(* Logix 5000 project; controller TFF vendor 1 type 14 code 107 rev 33.11; software revision 33.04; part 3 of 38 *)

        [4,3].ScaledMax := 100.0, [4,4].Tag := 'PCV012', [4,4].RawMax := 27648, [4,4].ScaledMax := 100.0, [4,5].Tag := 'SPARE', [4,5].RawMax := 27648, [4,5].ScaledMax := 100.0, [4,6].Tag := 'SPARE', [4,6].RawValue := -6912, [4,6].RawMax := 27648, [4,6].ScaledValue := -25.0, [4,6].ScaledMax := 100.0, [4,7].Tag := 'SPARE', [4,7].RawMax := 27648, [4,7].ScaledMax := 100.0, [4,8].Tag := 'AO#1', [4,8].RawMax := 2047, [4,8].ScaledMax := 100.0, [4,8].EnableCfg := 1, [4,9].Tag := 'AO#2', [4,9].RawMax := 2047, [4,9].ScaledMax := 100.0, [4,9].EnableCfg := 1, [4,10].Tag := 'AO#3', [4,10].RawMax := 2047, [4,10].ScaledMax := 100.0, [4,10].EnableCfg := 1, [4,11].Tag := 'AO#4', [4,11].RawMax := 2047, [4,11].ScaledMax := 100.0, [4,11].EnableCfg := 1, [5,0].Tag := 'SIC001', [5,0].RawMax := 27648, [5,0].ScaledMax := 100.0, [5,0].EnableCfg := 1, [5,1].Tag := 'SIC002', [5,1].RawMax := 27648, [5,1].ScaledMax := 100.0, [5,1].EnableCfg := 1, [5,2].Tag := 'PCV010', [5,2].RawMax := 2047, [5,2].ScaledMax := 100.0, [5,2].EnableCfg := 1, [5,3].Tag := 'PCV011', [5,3].RawMax := 27648, [5,3].ScaledMax := 100.0, [5,4].Tag := 'PCV012', [5,4].RawMax := 27648, [5,4].ScaledMax := 100.0, [5,5].Tag := 'SPARE', [5,5].RawMax := 27648, [5,5].ScaledMax := 100.0, [5,6].Tag := 'SPARE', [5,6].RawValue := -6912, [5,6].RawMax := 27648, [5,6].ScaledValue := -25.0, [5,6].ScaledMax := 100.0, [5,7].Tag := 'SPARE', [5,7].RawMax := 27648, [5,7].ScaledMax := 100.0,
        [5,8].Tag := 'AO#1', [5,8].RawMax := 2047, [5,8].ScaledMax := 100.0, [5,8].EnableCfg := 1, [5,9].Tag := 'AO#2', [5,9].RawMax := 2047, [5,9].ScaledMax := 100.0, [5,9].EnableCfg := 1, [5,10].Tag := 'AO#3', [5,10].RawMax := 2047, [5,10].ScaledMax := 100.0, [5,10].EnableCfg := 1, [5,11].Tag := 'AO#4', [5,11].RawMax := 2047, [5,11].ScaledMax := 100.0, [5,11].EnableCfg := 1);
   AnalogPoint : AnalogInput[50] := ([0].TagName := 'AI201B', [0].OutofRange := 1, [0].RawMin := 5529, [0].RawMax := 27648, [0].RawLowLimit := 5253, [0].RawHighLimit := 27924, [0].FilterActual := 1.0, [0].ScaledMax := 200.0, [0].CurrentValue := -49.993214, [0].RangeMax := 200.0, [0].RangeMaxSave := 200.0, [0].RealCfg := 1, [0].EnableCfg := 1, [0].OverrideCfg := 1, [0].EGU := 'mS/cm', [1].TagName := 'WI201', [1].OutofRange := 1, [1].Address := 1, [1].RawMin := 6553, [1].RawMax := 32767, [1].RawLowLimit := 6225, [1].RawHighLimit := 33095, [1].FilterActual := 1.0, [1].ScaledMax := 2000.0, [1].CurrentValue := -499.94724, [1].RangeMax := 2000.0, [1].RangeMaxSave := 2000.0, [1].RealCfg := 1, [1].EnableCfg := 1, [1].OverrideCfg := 1, [1].EGU := 'kg', [2].TagName := 'FI201', [2].OutofRange := 1, [2].Address := 2, [2].RawMin := 6553, [2].RawMax := 32767, [2].RawValue := 323, [2].RawLowLimit := 6225, [2].RawHighLimit := 33095, [2].FilteredRaw := 323, [2].FilterActual := 1.0, [2].ScaledMax := 100.0, [2].CurrentValue := -23.765926, [2].RangeMax := 100.0, [2].RangeMaxSave := 100.0, [2].RealCfg := 1, [2].EnableCfg := 1, [2].OverrideCfg := 1, [2].EGU := 'Lpm', [3].TagName := 'PCV101', [3].Address := 3, [3].RawMin := 6553, [3].RawMax := 32767, [3].RawValue := 12345, [3].RawLowLimit := 6225, [3].RawHighLimit := 33095, [3].FilteredRaw := 12345, [3].FilterActual := 1.0, [3].ScaledMax := 100.0, [3].CurrentValue := 0.059335444,
        [3].RangeMax := 100.0, [3].RangeMaxSave := 100.0, [3].EnableCfg := 1, [3].EGU := '%Clo', [4].TagName := 'PCV201', [4].Address := 4, [4].RawMin := 6553, [4].RawMax := 32767, [4].RawValue := 17653, [4].RawLowLimit := 6225, [4].RawHighLimit := 33095, [4].FilteredRaw := 17653, [4].FilterActual := 1.0, [4].ScaledMax := 100.0, [4].CurrentValue := 51.80897, [4].RangeMax := 100.0, [4].RangeMaxSave := 100.0, [4].EnableCfg := 1, [4].EGU := '%Opn', [5].TagName := 'PI001', [5].Address := 5, [5].RawMin := 6553, [5].RawMax := 32767, [5].RawValue := 32767, [5].RawLowLimit := 3276, [5].RawHighLimit := 33095, [5].FilteredRaw := 32767, [5].FilterActual := 1.0, [5].ScaledMax := 75.0, [5].CurrentValue := 75.0, [5].RangeMax := 75.0, [5].RangeMaxSave := 75.0, [5].RealCfg := 1, [5].EnableCfg := 1, [5].OverrideCfg := 1, [5].EGU := 'psi', [6].TagName := 'PI101', [6].Address := 6, [6].RawMin := 6553, [6].RawMax := 32767, [6].RawValue := 6576, [6].RawLowLimit := 3276, [6].RawHighLimit := 33095, [6].FilterUser := 50, [6].FilteredRaw := 6575, [6].FilterActual := 0.5, [6].ScaledMax := 75.0, [6].CurrentValue := 0.062943466, [6].RangeMax := 75.0, [6].RangeMaxSave := 75.0, [6].RealCfg := 1, [6].EnableCfg := 1, [6].OverrideCfg := 1, [6].EGU := 'psi', [7].TagName := 'PI201', [7].Address := 7, [7].RawMin := 6553, [7].RawMax := 32767, [7].RawValue := 6561, [7].RawLowLimit := 3276,
        [7].RawHighLimit := 33095, [7].FilteredRaw := 6561, [7].FilterActual := 1.0, [7].ScaledMax := 75.0, [7].CurrentValue := 0.022888534, [7].RangeMax := 75.0, [7].RangeMaxSave := 75.0, [7].RealCfg := 1, [7].EnableCfg := 1, [7].OverrideCfg := 1, [7].EGU := 'psi', [8].TagName := 'PI401', [8].Address := 8, [8].RawMin := 6553, [8].RawMax := 32767, [8].RawValue := 6563, [8].RawLowLimit := 3276, [8].RawHighLimit := 33095, [8].FilteredRaw := 6563, [8].FilterActual := 1.0, [8].ScaledMax := 75.0, [8].CurrentValue := 0.028610667, [8].RangeMax := 75.0, [8].RangeMaxSave := 75.0, [8].RealCfg := 1, [8].EnableCfg := 1, [8].OverrideCfg := 1, [8].EGU := 'psi', [9].TagName := 'AI202', [9].Address := 9, [9].RawMin := 5529, [9].RawMax := 27648, [9].RawLowLimit := 5253, [9].RawHighLimit := 27924, [9].FilterActual := 1.0, [9].ScaledMax := 14.0, [9].RangeMax := 14.0, [9].RangeMaxSave := 14.0, [9].EnableCfg := 1, [9].OverrideCfg := 1, [9].EGU := 'pH', [10].TagName := 'AI201A', [10].OutofRange := 1, [10].Address := 10, [10].RawMin := 5529, [10].RawMax := 27648, [10].RawLowLimit := 5253, [10].RawHighLimit := 27924, [10].FilterActual := 1.0, [10].ScaledMax := 120.0, [10].CurrentValue := -29.99593, [10].RangeMax := 120.0, [10].RangeMaxSave := 120.0, [10].RealCfg := 1, [10].EnableCfg := 1, [10].OverrideCfg := 1, [10].EGU := 'mS/cm', [11].TagName := 'AI203', [11].OutofRange := 1, [11].Address := 11,
        [11].RawMin := 5529, [11].RawMax := 27648, [11].RawLowLimit := 5253, [11].RawHighLimit := 27924, [11].FilterActual := 1.0, [11].ScaledMax := 2.0, [11].CurrentValue := -0.49993217, [11].RangeMax := 2.0, [11].RangeMaxSave := 2.0, [11].RealCfg := 1, [11].EnableCfg := 1, [11].OverrideCfg := 1, [11].EGU := 'AU', [12].TagName := 'AI204', [12].OutofRange := 1, [12].Address := 12, [12].RawMin := 5529, [12].RawMax := 27648, [12].RawLowLimit := 5253, [12].RawHighLimit := 27924, [12].FilterActual := 1.0, [12].ScaledMax := 2.0, [12].CurrentValue := -0.49993217, [12].RangeMax := 2.0, [12].RangeMaxSave := 2.0, [12].RealCfg := 1, [12].EnableCfg := 1, [12].OverrideCfg := 1, [12].EGU := 'AU', [13].TagName := 'TI101', [13].OutofRange := 1, [13].Address := 13, [13].RawMin := 5529, [13].RawMax := 27648, [13].RawLowLimit := 5253, [13].RawHighLimit := 27924, [13].FilterActual := 1.0, [13].ScaledMax := 100.0, [13].CurrentValue := -24.996607, [13].RangeMax := 100.0, [13].RangeMaxSave := 100.0, [13].RealCfg := 1, [13].EnableCfg := 1, [13].OverrideCfg := 1, [13].EGU := '$B0C', [14].TagName := 'MIX101', [14].Address := 14, [14].RawMax := 13824, [14].RawLowLimit := -138, [14].RawHighLimit := 13962, [14].FilterActual := 1.0, [14].ScaledMax := 100.0, [14].RangeMax := 100.0, [14].RangeMaxSave := 100.0, [14].RealCfg := 1, [14].EnableCfg := 1, [14].EGU := '%', [15].TagName := 'WI101', [15].Address := 15, [15].RawMax := 99999,
        [15].RawLowLimit := -1000, [15].RawHighLimit := 100999, [15].FilterActual := 1.0, [15].ScaledMax := 999.99, [15].CurrentValue := -127.832535, [15].EnableCfg := 1, [15].OverrideCfg := 1, [16].TagName := 'AI101', [16].Address := 16, [16].RawMin := 6553, [16].RawMax := 32767, [16].RawLowLimit := 6225, [16].RawHighLimit := 33095, [16].FilterActual := 1.0, [16].ScaledMax := 14.0, [16].RangeMax := 14.0, [16].RangeMaxSave := 14.0, [16].EnableCfg := 1, [16].OverrideCfg := 1, [16].EGU := 'pH', [17].TagName := 'AI104', [17].OutofRange := 1, [17].Address := 17, [17].RawMin := 5529, [17].RawMax := 27648, [17].RawLowLimit := 5253, [17].RawHighLimit := 27924, [17].FilterActual := 1.0, [17].ScaledMax := 200.0, [17].CurrentValue := -49.993214, [17].RangeMax := 200.0, [17].RangeMaxSave := 200.0, [17].RealCfg := 1, [17].OverrideCfg := 1, [17].EGU := 'mS/cm', [18].TagName := 'TCU101', [18].OutofRange := 1, [18].Address := 18, [18].RawMin := 5529, [18].RawMax := 27648, [18].RawLowLimit := 5253, [18].RawHighLimit := 27924, [18].FilterActual := 1.0, [18].ScaledMax := 100.0, [18].CurrentValue := -24.996607, [18].RangeMax := 100.0, [18].RangeMaxSave := 100.0, [18].RealCfg := 1, [18].OverrideCfg := 1, [18].EGU := '$B0C', [19].TagName := 'FI101', [19].Address := 19, [19].RawMin := 6553, [19].RawMax := 32767, [19].RawValue := 6555, [19].RawLowLimit := 6225, [19].RawHighLimit := 33095, [19].FilteredRaw := 6555, [19].FilterActual := 1.0, [19].ScaledMax := 100.0,
        [19].RangeMax := 100.0, [19].RangeMaxSave := 100.0, [19].EnableCfg := 1, [19].OverrideCfg := 1, [19].EGU := 'Lpm', [20].TagName := 'FI401', [20].Address := 20, [20].RawMin := 6553, [20].RawMax := 32767, [20].RawValue := 6550, [20].RawLowLimit := 6225, [20].RawHighLimit := 33095, [20].FilteredRaw := 6550, [20].FilterActual := 1.0, [20].ScaledMax := 100.0, [20].RangeMax := 100.0, [20].RangeMaxSave := 100.0, [20].EnableCfg := 1, [20].OverrideCfg := 1, [20].EGU := 'Lpm', [21].TagName := 'PI601', [21].OutofRange := 1, [21].Address := 21, [21].RawMin := 6553, [21].RawMax := 32767, [21].RawLowLimit := 3276, [21].RawHighLimit := 33095, [21].FilterActual := 1.0, [21].ScaledMax := 138.0, [21].CurrentValue := -34.497368, [21].RangeMax := 138.0, [21].RangeMaxSave := 138.0, [21].RealCfg := 1, [21].EnableCfg := 1, [21].OverrideCfg := 1, [21].EGU := 'mbar', [22].TagName := 'SPARE', [22].OutofRange := 1, [22].Address := 22, [22].RawMin := 5529, [22].RawMax := 27648, [22].RawLowLimit := 5253, [22].RawHighLimit := 27924, [22].FilterActual := 1.0, [22].ScaledMax := 100.0, [22].CurrentValue := -24.996607, [22].RangeMax := 100.0, [22].RangeMaxSave := 100.0, [22].RealCfg := 1, [22].EnableCfg := 1, [22].OverrideCfg := 1, [22].EGU := '$B0C', [23].TagName := 'SPARE', [24].TagName := 'SPARE', [25].TagName := 'SPARE', [26].TagName := 'SPARE', [27].TagName := 'SPARE', [28].TagName := 'AI1', [28].OutofRange := 1, [28].Address := 28,
        [28].RawMin := 6553, [28].RawMax := 32767, [28].RawLowLimit := 6225, [28].RawHighLimit := 33095, [28].FilterActual := 1.0, [28].ScaledMax := 100.0, [28].CurrentValue := -24.998093, [28].RangeMax := 100.0, [28].RangeMaxSave := 100.0, [28].RealCfg := 1, [28].EnableCfg := 1, [28].OverrideCfg := 1, [28].EGU := '%', [29].TagName := 'AI2', [29].OutofRange := 1, [29].Address := 29, [29].RawMin := 6553, [29].RawMax := 32767, [29].RawLowLimit := 6225, [29].RawHighLimit := 33095, [29].FilterActual := 1.0, [29].ScaledMax := 100.0, [29].CurrentValue := -24.998093, [29].RangeMax := 100.0, [29].RangeMaxSave := 100.0, [29].RealCfg := 1, [29].EnableCfg := 1, [29].OverrideCfg := 1, [29].EGU := '%', [30].TagName := 'AI3', [30].OutofRange := 1, [30].Address := 30, [30].RawMin := 6553, [30].RawMax := 32767, [30].RawLowLimit := 6225, [30].RawHighLimit := 33095, [30].FilterActual := 1.0, [30].ScaledMax := 100.0, [30].CurrentValue := -24.998093, [30].RangeMax := 100.0, [30].RangeMaxSave := 100.0, [30].RealCfg := 1, [30].EnableCfg := 1, [30].OverrideCfg := 1, [30].EGU := '%', [31].TagName := 'AI4', [31].OutofRange := 1, [31].Address := 31, [31].RawMin := 6553, [31].RawMax := 32767, [31].RawLowLimit := 6225, [31].RawHighLimit := 33095, [31].FilterActual := 1.0, [31].ScaledMax := 100.0, [31].CurrentValue := -24.998093, [31].RangeMax := 100.0, [31].RangeMaxSave := 100.0, [31].RealCfg := 1, [31].EnableCfg := 1, [31].OverrideCfg := 1,
        [31].EGU := '%', [40].TagName := 'DP', [40].Address := 40, [40].RawMin := 6553, [40].RawMax := 32767, [40].RawLowLimit := 6225, [40].RawHighLimit := 33095, [40].FilterActual := 1.0, [40].ScaledMax := 75.0, [40].CurrentValue := 74.93992, [40].RangeMax := 75.0, [40].RangeMaxSave := 75.0, [40].EnableCfg := 1, [40].OverrideCfg := 1, [40].EGU := 'psi', [41].TagName := 'TMP', [41].Address := 41, [41].RawMin := 6553, [41].RawMax := 32767, [41].RawLowLimit := 6225, [41].RawHighLimit := 33095, [41].FilterActual := 1.0, [41].ScaledMax := 75.0, [41].CurrentValue := 37.49857, [41].RangeMax := 75.0, [41].RangeMaxSave := 75.0, [41].EnableCfg := 1, [41].OverrideCfg := 1, [41].EGU := 'psi', [42].TagName := 'FI003', [42].Address := 42, [42].RawMin := 6553, [42].RawMax := 32767, [42].RawLowLimit := 6225, [42].RawHighLimit := 33095, [42].FilterActual := 1.0, [42].ScaledMax := 120.0, [42].RangeMax := 120.0, [42].RangeMaxSave := 120.0, [42].EnableCfg := 1, [42].OverrideCfg := 1, [42].EGU := 'Lpm', [43].Address := 43, [43].RawMin := 6553, [43].RawMax := 32767, [43].OverrideCfg := 1, [44].TagName := 'LI101', [44].Address := 44, [44].RawMin := 6553, [44].RawMax := 32767, [44].RawLowLimit := 6225, [44].RawHighLimit := 33095, [44].FilterActual := 1.0, [44].ScaledMax := 500.0, [44].CurrentValue := -126.566864, [44].RangeMax := 200.0, [44].RangeMaxSave := 200.0, [44].EnableCfg := 1, [44].OverrideCfg := 1, [45].TagName := 'NWP',
        [45].Address := 45, [45].RawMin := 6553, [45].RawMax := 32767, [45].RawLowLimit := 6225, [45].RawHighLimit := 33095, [45].FilterActual := 1.0, [45].ScaledMax := 999.0, [45].RangeMax := 999.0, [45].RangeMaxSave := 999.0, [45].EnableCfg := 1, [45].EGU := 'L/m$B2/', [46].TagName := 'PERM', [46].Address := 46, [46].RawMin := 6553, [46].RawMax := 32767, [46].RawLowLimit := 6225, [46].RawHighLimit := 33095, [46].FilterActual := 1.0, [46].ScaledMax := 999.0, [46].RangeMax := 999.0, [46].RangeMaxSave := 999.0, [46].EnableCfg := 1, [46].EGU := 'L/m$B2/');   // Analog Input Array
        [19]   // Retentate Flow
        [41]   // Trans-Membrane Pressure
        [28]   // Exchange AI#1
        [0]   // Filtrate Conductivity Cleaning
        [10]   // Filtrate Conductivity Process
        [11]   // Filtrate UV
        [12]   // Filtrate UV
        [13]   // Feed Tank Temperature
        [14]   // Mixer Speed
        [15]   // Feed Tank Weight
        [16]   // Feed Tank pH
        [17]   // Feed Tank Conductivity
        [18]   // TCU Temperature
        [1]   // External Filtrate Weight Scale
        [20]   // Transfer Pump Flow
        [21]   // Feed Tank Pressure
        [22]   // Filtrate Temperature
        [29]   // Exchange AI#2
        [30]   // Exchange AI#3
        [2]   // Filtrate Flow
        [31]   // Exchange AI#4
        [3]   // Retentate Pressure Control Valve Position
        [40]   // Differential Pressure
        [42]   // Feed Flow
        [44]   // Feed Tank volume
        [45]   // Normalized Water Permeability
        [46]   // Membrane Permeability
        [4]   // Filtrate Pressure Control Valve Position
        [5]   // Feed Pressure
        [6]   // Retentate Pressure
        [7]   // Filtrate Pressure
        [8]   // Transfer Pump Pressure
        [9]   // Filtrate pH
   AnalogPoint_Storage : AnalogInput[6,50] := ([0,0].TagName := 'PCV032', [0,0].OutofRange := 1, [0,0].RawMin := 6553, [0,0].RawMax := 32767, [0,0].RawValue := 1, [0,0].RawLowLimit := 6225, [0,0].RawHighLimit := 33095, [0,0].FilteredRaw := 1, [0,0].FilterActual := 1.0, [0,0].ScaledMax := 100.0, [0,0].CurrentValue := -24.994278, [0,0].RangeMax := 100.0, [0,0].RangeMaxSave := 100.0, [0,0].RealCfg := 1, [0,0].EnableCfg := 1, [0,0].OverrideCfg := 1, [0,1].TagName := 'AI201B', [0,1].OutofRange := 1, [0,1].Address := 1, [0,1].RawMin := 5529, [0,1].RawMax := 27648, [0,1].RawLowLimit := 5253, [0,1].RawHighLimit := 27924, [0,1].FilterActual := 1.0, [0,1].ScaledMax := 50.0, [0,1].CurrentValue := -12.498303, [0,1].RangeMax := 50.0, [0,1].RangeMaxSave := 50.0, [0,1].RealCfg := 1, [0,1].EnableCfg := 1, [0,1].OverrideCfg := 1, [0,2].TagName := 'AI201A', [0,2].OutofRange := 1, [0,2].Address := 2, [0,2].RawMin := 5529, [0,2].RawMax := 27648, [0,2].RawLowLimit := 5253, [0,2].RawHighLimit := 27924, [0,2].FilterActual := 1.0, [0,2].ScaledMax := 100.0, [0,2].CurrentValue := -24.996607, [0,2].RangeMax := 100.0, [0,2].RangeMaxSave := 100.0, [0,2].RealCfg := 1, [0,2].EnableCfg := 1, [0,2].OverrideCfg := 1, [0,3].TagName := 'AI202', [0,3].OutofRange := 1, [0,3].Address := 3, [0,3].RawMin := 5529, [0,3].RawMax := 27648, [0,3].RawLowLimit := 5253, [0,3].RawHighLimit := 27924, [0,3].FilterActual := 1.0, [0,3].ScaledMax := 14.0, [0,3].CurrentValue := -3.499525, [0,3].RangeMax := 14.0, [0,3].RangeMaxSave := 14.0, [0,3].RealCfg := 1, [0,3].EnableCfg := 1,
        [0,3].OverrideCfg := 1, [0,4].TagName := 'TI201', [0,4].OutofRange := 1, [0,4].Address := 4, [0,4].RawMin := 5529, [0,4].RawMax := 27648, [0,4].RawLowLimit := 5253, [0,4].RawHighLimit := 27924, [0,4].FilterActual := 1.0, [0,4].ScaledMax := 100.0, [0,4].CurrentValue := -24.996607, [0,4].RangeMax := 100.0, [0,4].RangeMaxSave := 100.0, [0,4].RealCfg := 1, [0,4].EnableCfg := 1, [0,4].OverrideCfg := 1, [0,5].TagName := 'AI203', [0,5].OutofRange := 1, [0,5].Address := 5, [0,5].RawMin := 5529, [0,5].RawMax := 27648, [0,5].RawLowLimit := 5253, [0,5].RawHighLimit := 27924, [0,5].FilterActual := 1.0, [0,5].ScaledMax := 2.0, [0,5].CurrentValue := -0.49993217, [0,5].RangeMax := 2.0, [0,5].RangeMaxSave := 2.0, [0,5].RealCfg := 1, [0,5].EnableCfg := 1, [0,5].OverrideCfg := 1, [0,6].TagName := 'AI204', [0,6].OutofRange := 1, [0,6].Address := 6, [0,6].RawMin := 5529, [0,6].RawMax := 27648, [0,6].RawLowLimit := 5253, [0,6].RawHighLimit := 27924, [0,6].FilterActual := 1.0, [0,6].ScaledMax := 2.0, [0,6].CurrentValue := -0.49993217, [0,6].RangeMax := 2.0, [0,6].RangeMaxSave := 2.0, [0,6].RealCfg := 1, [0,6].EnableCfg := 1, [0,6].OverrideCfg := 1, [0,7].TagName := 'AI102', [0,7].OutofRange := 1, [0,7].Address := 7, [0,7].RawMin := 5529, [0,7].RawMax := 27648, [0,7].RawLowLimit := 5253, [0,7].RawHighLimit := 27924, [0,7].FilterActual := 1.0, [0,7].ScaledMax := 100.0, [0,7].CurrentValue := -24.996607, [0,7].RangeMax := 100.0, [0,7].RangeMaxSave := 100.0, [0,7].RealCfg := 1, [0,7].EnableCfg := 1,
        [0,7].OverrideCfg := 1, [0,8].TagName := 'AI103', [0,8].OutofRange := 1, [0,8].Address := 8, [0,8].RawMin := 5529, [0,8].RawMax := 27648, [0,8].RawLowLimit := 5253, [0,8].RawHighLimit := 27924, [0,8].FilterActual := 1.0, [0,8].ScaledMax := 14.0, [0,8].CurrentValue := -3.499525, [0,8].RangeMax := 14.0, [0,8].RangeMaxSave := 14.0, [0,8].RealCfg := 1, [0,8].EnableCfg := 1, [0,8].OverrideCfg := 1, [0,9].TagName := 'PI003', [0,9].OutofRange := 1, [0,9].Address := 9, [0,9].RawMin := 6553, [0,9].RawMax := 32767, [0,9].RawLowLimit := 6225, [0,9].RawHighLimit := 33095, [0,9].FilterActual := 1.0, [0,9].ScaledMax := 6.0, [0,9].CurrentValue := -1.4998856, [0,9].RangeMax := 6.0, [0,9].RangeMaxSave := 6.0, [0,9].RealCfg := 1, [0,9].EnableCfg := 1, [0,9].OverrideCfg := 1, [0,10].TagName := 'FI001', [0,10].Address := 10, [0,10].RawMin := 5529, [0,10].RawMax := 27648, [0,10].RawLowLimit := 5253, [0,10].RawHighLimit := 27924, [0,10].FilterActual := 1.0, [0,10].ScaledMax := 22.0, [0,10].RangeMax := 22.0, [0,10].RangeMaxSave := 22.0, [0,10].EnableCfg := 1, [0,10].OverrideCfg := 1, [0,11].TagName := 'PI001', [0,11].OutofRange := 1, [0,11].Address := 11, [0,11].RawMin := 6553, [0,11].RawMax := 32767, [0,11].RawLowLimit := 6225, [0,11].RawHighLimit := 33095, [0,11].FilterActual := 1.0, [0,11].ScaledMax := 6.0, [0,11].CurrentValue := -1.4998856, [0,11].RangeMax := 6.0, [0,11].RangeMaxSave := 6.0, [0,11].RealCfg := 1, [0,11].EnableCfg := 1, [0,11].OverrideCfg := 1, [0,12].TagName := 'FI002', [0,12].Address := 12,
        [0,12].RawMin := 5529, [0,12].RawMax := 27648, [0,12].RawLowLimit := 5253, [0,12].RawHighLimit := 27924, [0,12].FilterActual := 1.0, [0,12].ScaledMax := 22.0, [0,12].RangeMax := 22.0, [0,12].RangeMaxSave := 22.0, [0,12].EnableCfg := 1, [0,12].OverrideCfg := 1, [0,13].TagName := 'PI002', [0,13].OutofRange := 1, [0,13].Address := 13, [0,13].RawMin := 6553, [0,13].RawMax := 32767, [0,13].RawLowLimit := 6225, [0,13].RawHighLimit := 33095, [0,13].FilterActual := 1.0, [0,13].ScaledMax := 6.0, [0,13].CurrentValue := -1.4998856, [0,13].RangeMax := 6.0, [0,13].RangeMaxSave := 6.0, [0,13].RealCfg := 1, [0,13].EnableCfg := 1, [0,13].OverrideCfg := 1, [0,14].OutofRange := 1, [0,14].Address := 14, [0,14].RawMin := 5529, [0,14].RawMax := 27648, [0,14].RawLowLimit := 5253, [0,14].RawHighLimit := 27924, [0,14].FilterActual := 1.0, [0,14].ScaledMax := 14.0, [0,14].RangeMax := 14.0, [0,14].RangeMaxSave := 14.0, [0,14].RealCfg := 1, [0,14].OverrideCfg := 1, [0,15].OutofRange := 1, [0,15].Address := 15, [0,15].RawMin := 5529, [0,15].RawMax := 27648, [0,15].RawLowLimit := 5253, [0,15].RawHighLimit := 27924, [0,15].FilterActual := 1.0, [0,15].ScaledMax := 2.0, [0,15].CurrentValue := -0.49993217, [0,15].RangeMax := 2.0, [0,15].RangeMaxSave := 2.0, [0,15].RealCfg := 1, [0,15].OverrideCfg := 1, [0,16].OutofRange := 1, [0,16].Address := 16, [0,16].RawMin := 5529, [0,16].RawMax := 27648, [0,16].RawLowLimit := 5253, [0,16].RawHighLimit := 27924, [0,16].FilterActual := 1.0, [0,16].ScaledMax := 2.0, [0,16].CurrentValue := -0.49993217, [0,16].RangeMax := 2.0,
        [0,16].RangeMaxSave := 2.0, [0,16].RealCfg := 1, [0,16].OverrideCfg := 1, [0,17].OutofRange := 1, [0,17].Address := 17, [0,17].RawMin := 5529, [0,17].RawMax := 27648, [0,17].RawLowLimit := 5253, [0,17].RawHighLimit := 27924, [0,17].FilterActual := 1.0, [0,17].ScaledMin := -1.0, [0,17].ScaledMax := 5.0, [0,17].CurrentValue := -2.4997964, [0,17].RangeMin := -1.0, [0,17].RangeMax := 5.0, [0,17].RangeMinSave := -1.0, [0,17].RangeMaxSave := 5.0, [0,17].RealCfg := 1, [0,17].OverrideCfg := 1, [0,18].OutofRange := 1, [0,18].Address := 18, [0,18].RawMin := 5529, [0,18].RawMax := 27648, [0,18].RawLowLimit := 5253, [0,18].RawHighLimit := 27924, [0,18].FilterActual := 1.0, [0,18].ScaledMin := -1.0, [0,18].ScaledMax := 5.0, [0,18].CurrentValue := -2.4997964, [0,18].RangeMin := -1.0, [0,18].RangeMax := 5.0, [0,18].RangeMinSave := -1.0, [0,18].RangeMaxSave := 5.0, [0,18].RealCfg := 1, [0,18].OverrideCfg := 1, [0,19].OutofRange := 1, [0,19].Address := 19, [0,19].RawMin := 5529, [0,19].RawMax := 27648, [0,19].RawLowLimit := 5253, [0,19].RawHighLimit := 27924, [0,19].FilterActual := 1.0, [0,19].ScaledMin := -1.0, [0,19].ScaledMax := 5.0, [0,19].CurrentValue := -2.4997964, [0,19].RangeMin := -1.0, [0,19].RangeMax := 5.0, [0,19].RangeMinSave := -1.0, [0,19].RangeMaxSave := 5.0, [0,19].RealCfg := 1, [0,19].OverrideCfg := 1, [0,20].OutofRange := 1, [0,20].Address := 20, [0,20].RawMin := 5529, [0,20].RawMax := 27648, [0,20].RawLowLimit := 5253, [0,20].RawHighLimit := 27924, [0,20].FilterActual := 1.0, [0,20].ScaledMax := 100.0, [0,20].CurrentValue := -24.996607,
        [0,20].RangeMax := 100.0, [0,20].RangeMaxSave := 100.0, [0,20].RealCfg := 1, [0,20].OverrideCfg := 1, [0,21].OutofRange := 1, [0,21].Address := 21, [0,21].RawMin := 5529, [0,21].RawMax := 27648, [0,21].RawLowLimit := 5253, [0,21].RawHighLimit := 27924, [0,21].FilterActual := 1.0, [0,21].ScaledMax := 100.0, [0,21].CurrentValue := -24.996607, [0,21].RangeMax := 100.0, [0,21].RangeMaxSave := 100.0, [0,21].RealCfg := 1, [0,21].OverrideCfg := 1, [0,22].TagName := 'SPARE', [0,22].Address := 22, [0,22].RawMin := 5529, [0,22].RawMax := 27648, [0,22].RealCfg := 1, [0,22].OverrideCfg := 1, [0,23].TagName := 'SPARE', [0,23].Address := 23, [0,23].RawMin := 5529, [0,23].RawMax := 27648, [0,23].RealCfg := 1, [0,23].OverrideCfg := 1, [0,24].TagName := 'SPARE', [0,24].Address := 24, [0,24].RawMin := 5529, [0,24].RawMax := 27648, [0,24].RealCfg := 1, [0,24].OverrideCfg := 1, [0,25].TagName := 'SPARE', [0,25].Address := 25, [0,25].RawMin := 5529, [0,25].RawMax := 27648, [0,25].RealCfg := 1, [0,25].OverrideCfg := 1, [0,26].TagName := 'SPARE', [0,26].Address := 26, [0,26].RawMin := 5529, [0,26].RawMax := 27648, [0,26].RealCfg := 1, [0,26].OverrideCfg := 1, [0,27].TagName := 'SPARE', [0,27].Address := 27, [0,27].RawMin := 5529, [0,27].RawMax := 27648, [0,27].RealCfg := 1, [0,27].OverrideCfg := 1, [0,28].TagName := 'AI#1', [0,28].OutofRange := 1, [0,28].Address := 28, [0,28].RawMin := 6553, [0,28].RawMax := 32767, [0,28].RawLowLimit := 6225, [0,28].RawHighLimit := 33095,
        [0,28].FilterActual := 1.0, [0,28].ScaledMax := 100.0, [0,28].CurrentValue := -24.998093, [0,28].RangeMax := 100.0, [0,28].RangeMaxSave := 100.0, [0,28].RealCfg := 1, [0,28].EnableCfg := 1, [0,28].OverrideCfg := 1, [0,29].TagName := 'AI#2', [0,29].OutofRange := 1, [0,29].Address := 29, [0,29].RawMin := 6553, [0,29].RawMax := 32767, [0,29].RawLowLimit := 6225, [0,29].RawHighLimit := 33095, [0,29].FilterActual := 1.0, [0,29].ScaledMax := 100.0, [0,29].CurrentValue := -24.998093, [0,29].RangeMax := 100.0, [0,29].RangeMaxSave := 100.0, [0,29].RealCfg := 1, [0,29].EnableCfg := 1, [0,29].OverrideCfg := 1, [0,30].TagName := 'AI#3', [0,30].OutofRange := 1, [0,30].Address := 30, [0,30].RawMin := 6553, [0,30].RawMax := 32767, [0,30].RawValue := 49, [0,30].RawLowLimit := 6225, [0,30].RawHighLimit := 33095, [0,30].FilteredRaw := 49, [0,30].FilterActual := 1.0, [0,30].ScaledMax := 100.0, [0,30].CurrentValue := -24.811169, [0,30].RangeMax := 100.0, [0,30].RangeMaxSave := 100.0, [0,30].RealCfg := 1, [0,30].EnableCfg := 1, [0,30].OverrideCfg := 1, [0,31].TagName := 'AI#4', [0,31].OutofRange := 1, [0,31].Address := 31, [0,31].RawMin := 6553, [0,31].RawMax := 32767, [0,31].RawValue := 48, [0,31].RawLowLimit := 6225, [0,31].RawHighLimit := 33095, [0,31].FilteredRaw := 48, [0,31].FilterActual := 1.0, [0,31].ScaledMax := 100.0, [0,31].CurrentValue := -24.814985, [0,31].RangeMax := 100.0, [0,31].RangeMaxSave := 100.0, [0,31].RealCfg := 1, [0,31].EnableCfg := 1, [0,31].OverrideCfg := 1, [0,40].TagName := 'FI003', [0,40].Address := 40, [0,40].RawMin := 5529,
        [0,40].RawMax := 27648, [0,40].RawLowLimit := 5253, [0,40].RawHighLimit := 27924, [0,40].FilterActual := 1.0, [0,40].ScaledMax := 44.0, [0,40].RangeMax := 44.0, [0,40].RangeMaxSave := 44.0, [0,40].EnableCfg := 1, [0,40].OverrideCfg := 1, [0,41].TagName := 'LV003', [0,41].Address := 41, [0,41].RawMin := 6553, [0,41].RawMax := 32767, [0,41].RawLowLimit := 6225, [0,41].RawHighLimit := 33095, [0,41].FilterActual := 1.0, [0,41].ScaledMax := 9999.0, [0,41].RangeMax := 9999.0, [0,41].RangeMaxSave := 9999.0, [0,41].EnableCfg := 1, [0,41].OverrideCfg := 1, [0,42].TagName := 'LV001', [0,42].Address := 42, [0,42].RawMin := 6553, [0,42].RawMax := 32767, [0,42].RawLowLimit := 6225, [0,42].RawHighLimit := 33095, [0,42].FilterActual := 1.0, [0,42].ScaledMax := 9999.0, [0,42].RangeMax := 9999.0, [0,42].RangeMaxSave := 9999.0, [0,42].EnableCfg := 1, [0,42].OverrideCfg := 1, [0,43].TagName := 'LV002', [0,43].Address := 43, [0,43].RawMin := 6553, [0,43].RawMax := 32767, [0,43].RawLowLimit := 6225, [0,43].RawHighLimit := 33095, [0,43].FilterActual := 1.0, [0,43].ScaledMax := 9999.0, [0,43].RangeMax := 9999.0, [0,43].RangeMaxSave := 9999.0, [0,43].EnableCfg := 1, [0,43].OverrideCfg := 1, [0,44].Address := 44, [0,44].RawMin := 6553, [0,44].RawMax := 32767, [0,44].RawLowLimit := 6225, [0,44].RawHighLimit := 33095, [0,44].FilterActual := 1.0, [0,44].ScaledMax := 99999.0, [0,44].RangeMax := 99999.0, [0,44].RangeMaxSave := 99999.0, [0,45].Address := 42, [0,45].RawMin := 6553, [0,45].RawMax := 32767, [0,45].RawLowLimit := 6225, [0,45].RawHighLimit := 33095, [0,45].FilterActual := 1.0,
        [0,45].ScaledMin := -1.0, [0,45].ScaledMax := 5.0, [0,45].RangeMin := -1.0, [0,45].RangeMax := 5.0, [0,45].RangeMinSave := -1.0, [0,45].RangeMaxSave := 5.0, [0,45].OverrideCfg := 1, [1,0].TagName := 'PCV032', [1,0].OutofRange := 1, [1,0].RawMin := 6553, [1,0].RawMax := 32767, [1,0].RawValue := 1, [1,0].RawLowLimit := 6225, [1,0].RawHighLimit := 33095, [1,0].FilteredRaw := 1, [1,0].FilterActual := 1.0, [1,0].ScaledMax := 100.0, [1,0].CurrentValue := -24.994278, [1,0].RangeMax := 100.0, [1,0].RangeMaxSave := 100.0, [1,0].RealCfg := 1, [1,0].EnableCfg := 1, [1,0].OverrideCfg := 1, [1,1].TagName := 'AI201B', [1,1].OutofRange := 1, [1,1].Address := 1, [1,1].RawMin := 5529, [1,1].RawMax := 27648, [1,1].RawLowLimit := 5253, [1,1].RawHighLimit := 27924, [1,1].FilterActual := 1.0, [1,1].ScaledMax := 50.0, [1,1].CurrentValue := -12.498303, [1,1].RangeMax := 50.0, [1,1].RangeMaxSave := 50.0, [1,1].RealCfg := 1, [1,1].EnableCfg := 1, [1,1].OverrideCfg := 1, [1,2].TagName := 'AI201A', [1,2].OutofRange := 1, [1,2].Address := 2, [1,2].RawMin := 5529, [1,2].RawMax := 27648, [1,2].RawLowLimit := 5253, [1,2].RawHighLimit := 27924, [1,2].FilterActual := 1.0, [1,2].ScaledMax := 100.0, [1,2].CurrentValue := -24.996607, [1,2].RangeMax := 100.0, [1,2].RangeMaxSave := 100.0, [1,2].RealCfg := 1, [1,2].EnableCfg := 1, [1,2].OverrideCfg := 1, [1,3].TagName := 'AI202', [1,3].OutofRange := 1, [1,3].Address := 3, [1,3].RawMin := 5529, [1,3].RawMax := 27648, [1,3].RawLowLimit := 5253, [1,3].RawHighLimit := 27924,
        [1,3].FilterActual := 1.0, [1,3].ScaledMax := 14.0, [1,3].CurrentValue := -3.499525, [1,3].RangeMax := 14.0, [1,3].RangeMaxSave := 14.0, [1,3].RealCfg := 1, [1,3].EnableCfg := 1, [1,3].OverrideCfg := 1, [1,4].TagName := 'TI201', [1,4].OutofRange := 1, [1,4].Address := 4, [1,4].RawMin := 5529, [1,4].RawMax := 27648, [1,4].RawLowLimit := 5253, [1,4].RawHighLimit := 27924, [1,4].FilterActual := 1.0, [1,4].ScaledMax := 100.0, [1,4].CurrentValue := -24.996607, [1,4].RangeMax := 100.0, [1,4].RangeMaxSave := 100.0, [1,4].RealCfg := 1, [1,4].EnableCfg := 1, [1,4].OverrideCfg := 1, [1,5].TagName := 'AI203', [1,5].OutofRange := 1, [1,5].Address := 5, [1,5].RawMin := 5529, [1,5].RawMax := 27648, [1,5].RawLowLimit := 5253, [1,5].RawHighLimit := 27924, [1,5].FilterActual := 1.0, [1,5].ScaledMax := 2.0, [1,5].CurrentValue := -0.49993217, [1,5].RangeMax := 2.0, [1,5].RangeMaxSave := 2.0, [1,5].RealCfg := 1, [1,5].EnableCfg := 1, [1,5].OverrideCfg := 1, [1,6].TagName := 'AI204', [1,6].OutofRange := 1, [1,6].Address := 6, [1,6].RawMin := 5529, [1,6].RawMax := 27648, [1,6].RawLowLimit := 5253, [1,6].RawHighLimit := 27924, [1,6].FilterActual := 1.0, [1,6].ScaledMax := 2.0, [1,6].CurrentValue := -0.49993217, [1,6].RangeMax := 2.0, [1,6].RangeMaxSave := 2.0, [1,6].RealCfg := 1, [1,6].EnableCfg := 1, [1,6].OverrideCfg := 1, [1,7].TagName := 'AI102', [1,7].OutofRange := 1, [1,7].Address := 7, [1,7].RawMin := 5529, [1,7].RawMax := 27648, [1,7].RawLowLimit := 5253, [1,7].RawHighLimit := 27924,
        [1,7].FilterActual := 1.0, [1,7].ScaledMax := 100.0, [1,7].CurrentValue := -24.996607, [1,7].RangeMax := 100.0, [1,7].RangeMaxSave := 100.0, [1,7].RealCfg := 1, [1,7].EnableCfg := 1, [1,7].OverrideCfg := 1, [1,8].TagName := 'AI103', [1,8].OutofRange := 1, [1,8].Address := 8, [1,8].RawMin := 5529, [1,8].RawMax := 27648, [1,8].RawLowLimit := 5253, [1,8].RawHighLimit := 27924, [1,8].FilterActual := 1.0, [1,8].ScaledMax := 14.0, [1,8].CurrentValue := -3.499525, [1,8].RangeMax := 14.0, [1,8].RangeMaxSave := 14.0, [1,8].RealCfg := 1, [1,8].EnableCfg := 1, [1,8].OverrideCfg := 1, [1,9].TagName := 'PI003', [1,9].OutofRange := 1, [1,9].Address := 9, [1,9].RawMin := 6553, [1,9].RawMax := 32767, [1,9].RawLowLimit := 6225, [1,9].RawHighLimit := 33095, [1,9].FilterActual := 1.0, [1,9].ScaledMax := 6.0, [1,9].CurrentValue := -1.4998856, [1,9].RangeMax := 6.0, [1,9].RangeMaxSave := 6.0, [1,9].RealCfg := 1, [1,9].EnableCfg := 1, [1,9].OverrideCfg := 1, [1,10].TagName := 'FI001', [1,10].Address := 10, [1,10].RawMin := 5529, [1,10].RawMax := 27648, [1,10].RawLowLimit := 5253, [1,10].RawHighLimit := 27924, [1,10].FilterActual := 1.0, [1,10].ScaledMax := 22.0, [1,10].RangeMax := 22.0, [1,10].RangeMaxSave := 22.0, [1,10].EnableCfg := 1, [1,10].OverrideCfg := 1, [1,11].TagName := 'PI001', [1,11].OutofRange := 1, [1,11].Address := 11, [1,11].RawMin := 6553, [1,11].RawMax := 32767, [1,11].RawLowLimit := 6225, [1,11].RawHighLimit := 33095, [1,11].FilterActual := 1.0, [1,11].ScaledMax := 6.0, [1,11].CurrentValue := -1.4998856,
        [1,11].RangeMax := 6.0, [1,11].RangeMaxSave := 6.0, [1,11].RealCfg := 1, [1,11].EnableCfg := 1, [1,11].OverrideCfg := 1, [1,12].TagName := 'FI002', [1,12].Address := 12, [1,12].RawMin := 5529, [1,12].RawMax := 27648, [1,12].RawLowLimit := 5253, [1,12].RawHighLimit := 27924, [1,12].FilterActual := 1.0, [1,12].ScaledMax := 22.0, [1,12].RangeMax := 22.0, [1,12].RangeMaxSave := 22.0, [1,12].EnableCfg := 1, [1,12].OverrideCfg := 1, [1,13].TagName := 'PI002', [1,13].OutofRange := 1, [1,13].Address := 13, [1,13].RawMin := 6553, [1,13].RawMax := 32767, [1,13].RawLowLimit := 6225, [1,13].RawHighLimit := 33095, [1,13].FilterActual := 1.0, [1,13].ScaledMax := 6.0, [1,13].CurrentValue := -1.4998856, [1,13].RangeMax := 6.0, [1,13].RangeMaxSave := 6.0, [1,13].RealCfg := 1, [1,13].EnableCfg := 1, [1,13].OverrideCfg := 1, [1,14].OutofRange := 1, [1,14].Address := 14, [1,14].RawMin := 5529, [1,14].RawMax := 27648, [1,14].RawLowLimit := 5253, [1,14].RawHighLimit := 27924, [1,14].FilterActual := 1.0, [1,14].ScaledMax := 14.0, [1,14].RangeMax := 14.0, [1,14].RangeMaxSave := 14.0, [1,14].RealCfg := 1, [1,14].OverrideCfg := 1, [1,15].OutofRange := 1, [1,15].Address := 15, [1,15].RawMin := 5529, [1,15].RawMax := 27648, [1,15].RawLowLimit := 5253, [1,15].RawHighLimit := 27924, [1,15].FilterActual := 1.0, [1,15].ScaledMax := 2.0, [1,15].CurrentValue := -0.49993217, [1,15].RangeMax := 2.0, [1,15].RangeMaxSave := 2.0, [1,15].RealCfg := 1, [1,15].OverrideCfg := 1, [1,16].OutofRange := 1, [1,16].Address := 16, [1,16].RawMin := 5529,
        [1,16].RawMax := 27648, [1,16].RawLowLimit := 5253, [1,16].RawHighLimit := 27924, [1,16].FilterActual := 1.0, [1,16].ScaledMax := 2.0, [1,16].CurrentValue := -0.49993217, [1,16].RangeMax := 2.0, [1,16].RangeMaxSave := 2.0, [1,16].RealCfg := 1, [1,16].OverrideCfg := 1, [1,17].OutofRange := 1, [1,17].Address := 17, [1,17].RawMin := 5529, [1,17].RawMax := 27648, [1,17].RawLowLimit := 5253, [1,17].RawHighLimit := 27924, [1,17].FilterActual := 1.0, [1,17].ScaledMin := -1.0, [1,17].ScaledMax := 5.0, [1,17].CurrentValue := -2.4997964, [1,17].RangeMin := -1.0, [1,17].RangeMax := 5.0, [1,17].RangeMinSave := -1.0, [1,17].RangeMaxSave := 5.0, [1,17].RealCfg := 1, [1,17].OverrideCfg := 1, [1,18].OutofRange := 1, [1,18].Address := 18, [1,18].RawMin := 5529, [1,18].RawMax := 27648, [1,18].RawLowLimit := 5253, [1,18].RawHighLimit := 27924, [1,18].FilterActual := 1.0, [1,18].ScaledMin := -1.0, [1,18].ScaledMax := 5.0, [1,18].CurrentValue := -2.4997964, [1,18].RangeMin := -1.0, [1,18].RangeMax := 5.0, [1,18].RangeMinSave := -1.0, [1,18].RangeMaxSave := 5.0, [1,18].RealCfg := 1, [1,18].OverrideCfg := 1, [1,19].OutofRange := 1, [1,19].Address := 19, [1,19].RawMin := 5529, [1,19].RawMax := 27648, [1,19].RawLowLimit := 5253, [1,19].RawHighLimit := 27924, [1,19].FilterActual := 1.0, [1,19].ScaledMin := -1.0, [1,19].ScaledMax := 5.0, [1,19].CurrentValue := -2.4997964, [1,19].RangeMin := -1.0, [1,19].RangeMax := 5.0, [1,19].RangeMinSave := -1.0, [1,19].RangeMaxSave := 5.0, [1,19].RealCfg := 1, [1,19].OverrideCfg := 1, [1,20].OutofRange := 1, [1,20].Address := 20,
        [1,20].RawMin := 5529, [1,20].RawMax := 27648, [1,20].RawLowLimit := 5253, [1,20].RawHighLimit := 27924, [1,20].FilterActual := 1.0, [1,20].ScaledMax := 100.0, [1,20].CurrentValue := -24.996607, [1,20].RangeMax := 100.0, [1,20].RangeMaxSave := 100.0, [1,20].RealCfg := 1, [1,20].OverrideCfg := 1, [1,21].OutofRange := 1, [1,21].Address := 21, [1,21].RawMin := 5529, [1,21].RawMax := 27648, [1,21].RawLowLimit := 5253, [1,21].RawHighLimit := 27924, [1,21].FilterActual := 1.0, [1,21].ScaledMax := 100.0, [1,21].CurrentValue := -24.996607, [1,21].RangeMax := 100.0, [1,21].RangeMaxSave := 100.0, [1,21].RealCfg := 1, [1,21].OverrideCfg := 1, [1,22].TagName := 'SPARE', [1,22].Address := 22, [1,22].RawMin := 5529, [1,22].RawMax := 27648, [1,22].RealCfg := 1, [1,22].OverrideCfg := 1, [1,23].TagName := 'SPARE', [1,23].Address := 23, [1,23].RawMin := 5529, [1,23].RawMax := 27648, [1,23].RealCfg := 1, [1,23].OverrideCfg := 1, [1,24].TagName := 'SPARE', [1,24].Address := 24, [1,24].RawMin := 5529, [1,24].RawMax := 27648, [1,24].RealCfg := 1, [1,24].OverrideCfg := 1, [1,25].TagName := 'SPARE', [1,25].Address := 25, [1,25].RawMin := 5529, [1,25].RawMax := 27648, [1,25].RealCfg := 1, [1,25].OverrideCfg := 1, [1,26].TagName := 'SPARE', [1,26].Address := 26, [1,26].RawMin := 5529, [1,26].RawMax := 27648, [1,26].RealCfg := 1, [1,26].OverrideCfg := 1, [1,27].TagName := 'SPARE', [1,27].Address := 27, [1,27].RawMin := 5529, [1,27].RawMax := 27648, [1,27].RealCfg := 1, [1,27].OverrideCfg := 1,
        [1,28].TagName := 'AI#1', [1,28].OutofRange := 1, [1,28].Address := 28, [1,28].RawMin := 6553, [1,28].RawMax := 32767, [1,28].RawLowLimit := 6225, [1,28].RawHighLimit := 33095, [1,28].FilterActual := 1.0, [1,28].ScaledMax := 100.0, [1,28].CurrentValue := -24.998093, [1,28].RangeMax := 100.0, [1,28].RangeMaxSave := 100.0, [1,28].RealCfg := 1, [1,28].EnableCfg := 1, [1,28].OverrideCfg := 1, [1,29].TagName := 'AI#2', [1,29].OutofRange := 1, [1,29].Address := 29, [1,29].RawMin := 6553, [1,29].RawMax := 32767, [1,29].RawLowLimit := 6225, [1,29].RawHighLimit := 33095, [1,29].FilterActual := 1.0, [1,29].ScaledMax := 100.0, [1,29].CurrentValue := -24.998093, [1,29].RangeMax := 100.0, [1,29].RangeMaxSave := 100.0, [1,29].RealCfg := 1, [1,29].EnableCfg := 1, [1,29].OverrideCfg := 1, [1,30].TagName := 'AI#3', [1,30].OutofRange := 1, [1,30].Address := 30, [1,30].RawMin := 6553, [1,30].RawMax := 32767, [1,30].RawValue := 49, [1,30].RawLowLimit := 6225, [1,30].RawHighLimit := 33095, [1,30].FilteredRaw := 49, [1,30].FilterActual := 1.0, [1,30].ScaledMax := 100.0, [1,30].CurrentValue := -24.811169, [1,30].RangeMax := 100.0, [1,30].RangeMaxSave := 100.0, [1,30].RealCfg := 1, [1,30].EnableCfg := 1, [1,30].OverrideCfg := 1, [1,31].TagName := 'AI#4', [1,31].OutofRange := 1, [1,31].Address := 31, [1,31].RawMin := 6553, [1,31].RawMax := 32767, [1,31].RawValue := 48, [1,31].RawLowLimit := 6225, [1,31].RawHighLimit := 33095, [1,31].FilteredRaw := 48, [1,31].FilterActual := 1.0, [1,31].ScaledMax := 100.0, [1,31].CurrentValue := -24.814985, [1,31].RangeMax := 100.0,
        [1,31].RangeMaxSave := 100.0, [1,31].RealCfg := 1, [1,31].EnableCfg := 1, [1,31].OverrideCfg := 1, [1,40].TagName := 'FI003', [1,40].Address := 40, [1,40].RawMin := 5529, [1,40].RawMax := 27648, [1,40].RawLowLimit := 5253, [1,40].RawHighLimit := 27924, [1,40].FilterActual := 1.0, [1,40].ScaledMax := 44.0, [1,40].RangeMax := 44.0, [1,40].RangeMaxSave := 44.0, [1,40].EnableCfg := 1, [1,40].OverrideCfg := 1, [1,41].TagName := 'LV003', [1,41].Address := 41, [1,41].RawMin := 6553, [1,41].RawMax := 32767, [1,41].RawLowLimit := 6225, [1,41].RawHighLimit := 33095, [1,41].FilterActual := 1.0, [1,41].ScaledMax := 9999.0, [1,41].RangeMax := 9999.0, [1,41].RangeMaxSave := 9999.0, [1,41].EnableCfg := 1, [1,41].OverrideCfg := 1, [1,42].TagName := 'LV001', [1,42].Address := 42, [1,42].RawMin := 6553, [1,42].RawMax := 32767, [1,42].RawLowLimit := 6225, [1,42].RawHighLimit := 33095, [1,42].FilterActual := 1.0, [1,42].ScaledMax := 9999.0, [1,42].RangeMax := 9999.0, [1,42].RangeMaxSave := 9999.0, [1,42].EnableCfg := 1, [1,42].OverrideCfg := 1, [1,43].TagName := 'LV002', [1,43].Address := 43, [1,43].RawMin := 6553, [1,43].RawMax := 32767, [1,43].RawLowLimit := 6225, [1,43].RawHighLimit := 33095, [1,43].FilterActual := 1.0, [1,43].ScaledMax := 9999.0, [1,43].RangeMax := 9999.0, [1,43].RangeMaxSave := 9999.0, [1,43].EnableCfg := 1, [1,43].OverrideCfg := 1, [1,44].Address := 44, [1,44].RawMin := 6553, [1,44].RawMax := 32767, [1,44].RawLowLimit := 6225, [1,44].RawHighLimit := 33095, [1,44].FilterActual := 1.0, [1,44].ScaledMax := 99999.0, [1,44].RangeMax := 99999.0,
        [1,44].RangeMaxSave := 99999.0, [1,45].Address := 42, [1,45].RawMin := 6553, [1,45].RawMax := 32767, [1,45].RawLowLimit := 6225, [1,45].RawHighLimit := 33095, [1,45].FilterActual := 1.0, [1,45].ScaledMin := -1.0, [1,45].ScaledMax := 5.0, [1,45].RangeMin := -1.0, [1,45].RangeMax := 5.0, [1,45].RangeMinSave := -1.0, [1,45].RangeMaxSave := 5.0, [1,45].OverrideCfg := 1, [2,0].TagName := 'PCV032', [2,0].OutofRange := 1, [2,0].RawMin := 6553, [2,0].RawMax := 32767, [2,0].RawValue := 1, [2,0].RawLowLimit := 6225, [2,0].RawHighLimit := 33095, [2,0].FilteredRaw := 1, [2,0].FilterActual := 1.0, [2,0].ScaledMax := 100.0, [2,0].CurrentValue := -24.994278, [2,0].RangeMax := 100.0, [2,0].RangeMaxSave := 100.0, [2,0].RealCfg := 1, [2,0].EnableCfg := 1, [2,0].OverrideCfg := 1, [2,1].TagName := 'AI201B', [2,1].OutofRange := 1, [2,1].Address := 1, [2,1].RawMin := 5529, [2,1].RawMax := 27648, [2,1].RawLowLimit := 5253, [2,1].RawHighLimit := 27924, [2,1].FilterActual := 1.0, [2,1].ScaledMax := 50.0, [2,1].CurrentValue := -12.498303, [2,1].RangeMax := 50.0, [2,1].RangeMaxSave := 50.0, [2,1].RealCfg := 1, [2,1].EnableCfg := 1, [2,1].OverrideCfg := 1, [2,2].TagName := 'AI201A', [2,2].OutofRange := 1, [2,2].Address := 2, [2,2].RawMin := 5529, [2,2].RawMax := 27648, [2,2].RawLowLimit := 5253, [2,2].RawHighLimit := 27924, [2,2].FilterActual := 1.0, [2,2].ScaledMax := 100.0, [2,2].CurrentValue := -24.996607, [2,2].RangeMax := 100.0, [2,2].RangeMaxSave := 100.0, [2,2].RealCfg := 1, [2,2].EnableCfg := 1, [2,2].OverrideCfg := 1,
        [2,3].TagName := 'AI202', [2,3].OutofRange := 1, [2,3].Address := 3, [2,3].RawMin := 5529, [2,3].RawMax := 27648, [2,3].RawLowLimit := 5253, [2,3].RawHighLimit := 27924, [2,3].FilterActual := 1.0, [2,3].ScaledMax := 14.0, [2,3].CurrentValue := -3.499525, [2,3].RangeMax := 14.0, [2,3].RangeMaxSave := 14.0, [2,3].RealCfg := 1, [2,3].EnableCfg := 1, [2,3].OverrideCfg := 1, [2,4].TagName := 'TI201', [2,4].OutofRange := 1, [2,4].Address := 4, [2,4].RawMin := 5529, [2,4].RawMax := 27648, [2,4].RawLowLimit := 5253, [2,4].RawHighLimit := 27924, [2,4].FilterActual := 1.0, [2,4].ScaledMax := 100.0, [2,4].CurrentValue := -24.996607, [2,4].RangeMax := 100.0, [2,4].RangeMaxSave := 100.0, [2,4].RealCfg := 1, [2,4].EnableCfg := 1, [2,4].OverrideCfg := 1, [2,5].TagName := 'AI203', [2,5].OutofRange := 1, [2,5].Address := 5, [2,5].RawMin := 5529, [2,5].RawMax := 27648, [2,5].RawLowLimit := 5253, [2,5].RawHighLimit := 27924, [2,5].FilterActual := 1.0, [2,5].ScaledMax := 2.0, [2,5].CurrentValue := -0.49993217, [2,5].RangeMax := 2.0, [2,5].RangeMaxSave := 2.0, [2,5].RealCfg := 1, [2,5].EnableCfg := 1, [2,5].OverrideCfg := 1, [2,6].TagName := 'AI204', [2,6].OutofRange := 1, [2,6].Address := 6, [2,6].RawMin := 5529, [2,6].RawMax := 27648, [2,6].RawLowLimit := 5253, [2,6].RawHighLimit := 27924, [2,6].FilterActual := 1.0, [2,6].ScaledMax := 2.0, [2,6].CurrentValue := -0.49993217, [2,6].RangeMax := 2.0, [2,6].RangeMaxSave := 2.0, [2,6].RealCfg := 1, [2,6].EnableCfg := 1, [2,6].OverrideCfg := 1,
        [2,7].TagName := 'AI102', [2,7].OutofRange := 1, [2,7].Address := 7, [2,7].RawMin := 5529, [2,7].RawMax := 27648, [2,7].RawLowLimit := 5253, [2,7].RawHighLimit := 27924, [2,7].FilterActual := 1.0, [2,7].ScaledMax := 100.0, [2,7].CurrentValue := -24.996607, [2,7].RangeMax := 100.0, [2,7].RangeMaxSave := 100.0, [2,7].RealCfg := 1, [2,7].EnableCfg := 1, [2,7].OverrideCfg := 1, [2,8].TagName := 'AI103', [2,8].OutofRange := 1, [2,8].Address := 8, [2,8].RawMin := 5529, [2,8].RawMax := 27648, [2,8].RawLowLimit := 5253, [2,8].RawHighLimit := 27924, [2,8].FilterActual := 1.0, [2,8].ScaledMax := 14.0, [2,8].CurrentValue := -3.499525, [2,8].RangeMax := 14.0, [2,8].RangeMaxSave := 14.0, [2,8].RealCfg := 1, [2,8].EnableCfg := 1, [2,8].OverrideCfg := 1, [2,9].TagName := 'PI003', [2,9].OutofRange := 1, [2,9].Address := 9, [2,9].RawMin := 6553, [2,9].RawMax := 32767, [2,9].RawLowLimit := 6225, [2,9].RawHighLimit := 33095, [2,9].FilterActual := 1.0, [2,9].ScaledMax := 6.0, [2,9].CurrentValue := -1.4998856, [2,9].RangeMax := 6.0, [2,9].RangeMaxSave := 6.0, [2,9].RealCfg := 1, [2,9].EnableCfg := 1, [2,9].OverrideCfg := 1, [2,10].TagName := 'FI001', [2,10].Address := 10, [2,10].RawMin := 5529, [2,10].RawMax := 27648, [2,10].RawLowLimit := 5253, [2,10].RawHighLimit := 27924, [2,10].FilterActual := 1.0, [2,10].ScaledMax := 22.0, [2,10].RangeMax := 22.0, [2,10].RangeMaxSave := 22.0, [2,10].EnableCfg := 1, [2,10].OverrideCfg := 1, [2,11].TagName := 'PI001', [2,11].OutofRange := 1, [2,11].Address := 11,
        [2,11].RawMin := 6553, [2,11].RawMax := 32767, [2,11].RawLowLimit := 6225, [2,11].RawHighLimit := 33095, [2,11].FilterActual := 1.0, [2,11].ScaledMax := 6.0, [2,11].CurrentValue := -1.4998856, [2,11].RangeMax := 6.0, [2,11].RangeMaxSave := 6.0, [2,11].RealCfg := 1, [2,11].EnableCfg := 1, [2,11].OverrideCfg := 1, [2,12].TagName := 'FI002', [2,12].Address := 12, [2,12].RawMin := 5529, [2,12].RawMax := 27648, [2,12].RawLowLimit := 5253, [2,12].RawHighLimit := 27924, [2,12].FilterActual := 1.0, [2,12].ScaledMax := 22.0, [2,12].RangeMax := 22.0, [2,12].RangeMaxSave := 22.0, [2,12].EnableCfg := 1, [2,12].OverrideCfg := 1, [2,13].TagName := 'PI002', [2,13].OutofRange := 1, [2,13].Address := 13, [2,13].RawMin := 6553, [2,13].RawMax := 32767, [2,13].RawLowLimit := 6225, [2,13].RawHighLimit := 33095, [2,13].FilterActual := 1.0, [2,13].ScaledMax := 6.0, [2,13].CurrentValue := -1.4998856, [2,13].RangeMax := 6.0, [2,13].RangeMaxSave := 6.0, [2,13].RealCfg := 1, [2,13].EnableCfg := 1, [2,13].OverrideCfg := 1, [2,14].OutofRange := 1, [2,14].Address := 14, [2,14].RawMin := 5529, [2,14].RawMax := 27648, [2,14].RawLowLimit := 5253, [2,14].RawHighLimit := 27924, [2,14].FilterActual := 1.0, [2,14].ScaledMax := 14.0, [2,14].RangeMax := 14.0, [2,14].RangeMaxSave := 14.0, [2,14].RealCfg := 1, [2,14].OverrideCfg := 1, [2,15].OutofRange := 1, [2,15].Address := 15, [2,15].RawMin := 5529, [2,15].RawMax := 27648, [2,15].RawLowLimit := 5253, [2,15].RawHighLimit := 27924, [2,15].FilterActual := 1.0, [2,15].ScaledMax := 2.0, [2,15].CurrentValue := -0.49993217,
        [2,15].RangeMax := 2.0, [2,15].RangeMaxSave := 2.0, [2,15].RealCfg := 1, [2,15].OverrideCfg := 1, [2,16].OutofRange := 1, [2,16].Address := 16, [2,16].RawMin := 5529, [2,16].RawMax := 27648, [2,16].RawLowLimit := 5253, [2,16].RawHighLimit := 27924, [2,16].FilterActual := 1.0, [2,16].ScaledMax := 2.0, [2,16].CurrentValue := -0.49993217, [2,16].RangeMax := 2.0, [2,16].RangeMaxSave := 2.0, [2,16].RealCfg := 1, [2,16].OverrideCfg := 1, [2,17].OutofRange := 1, [2,17].Address := 17, [2,17].RawMin := 5529, [2,17].RawMax := 27648, [2,17].RawLowLimit := 5253, [2,17].RawHighLimit := 27924, [2,17].FilterActual := 1.0, [2,17].ScaledMin := -1.0, [2,17].ScaledMax := 5.0, [2,17].CurrentValue := -2.4997964, [2,17].RangeMin := -1.0, [2,17].RangeMax := 5.0, [2,17].RangeMinSave := -1.0, [2,17].RangeMaxSave := 5.0, [2,17].RealCfg := 1, [2,17].OverrideCfg := 1, [2,18].OutofRange := 1, [2,18].Address := 18, [2,18].RawMin := 5529, [2,18].RawMax := 27648, [2,18].RawLowLimit := 5253, [2,18].RawHighLimit := 27924, [2,18].FilterActual := 1.0, [2,18].ScaledMin := -1.0, [2,18].ScaledMax := 5.0, [2,18].CurrentValue := -2.4997964, [2,18].RangeMin := -1.0, [2,18].RangeMax := 5.0, [2,18].RangeMinSave := -1.0, [2,18].RangeMaxSave := 5.0, [2,18].RealCfg := 1, [2,18].OverrideCfg := 1, [2,19].OutofRange := 1, [2,19].Address := 19, [2,19].RawMin := 5529, [2,19].RawMax := 27648, [2,19].RawLowLimit := 5253, [2,19].RawHighLimit := 27924, [2,19].FilterActual := 1.0, [2,19].ScaledMin := -1.0, [2,19].ScaledMax := 5.0, [2,19].CurrentValue := -2.4997964, [2,19].RangeMin := -1.0,
        [2,19].RangeMax := 5.0, [2,19].RangeMinSave := -1.0, [2,19].RangeMaxSave := 5.0, [2,19].RealCfg := 1, [2,19].OverrideCfg := 1, [2,20].OutofRange := 1, [2,20].Address := 20, [2,20].RawMin := 5529, [2,20].RawMax := 27648, [2,20].RawLowLimit := 5253, [2,20].RawHighLimit := 27924, [2,20].FilterActual := 1.0, [2,20].ScaledMax := 100.0, [2,20].CurrentValue := -24.996607, [2,20].RangeMax := 100.0, [2,20].RangeMaxSave := 100.0, [2,20].RealCfg := 1, [2,20].OverrideCfg := 1, [2,21].OutofRange := 1, [2,21].Address := 21, [2,21].RawMin := 5529, [2,21].RawMax := 27648, [2,21].RawLowLimit := 5253, [2,21].RawHighLimit := 27924, [2,21].FilterActual := 1.0, [2,21].ScaledMax := 100.0, [2,21].CurrentValue := -24.996607, [2,21].RangeMax := 100.0, [2,21].RangeMaxSave := 100.0, [2,21].RealCfg := 1, [2,21].OverrideCfg := 1, [2,22].TagName := 'SPARE', [2,22].Address := 22, [2,22].RawMin := 5529, [2,22].RawMax := 27648, [2,22].RealCfg := 1, [2,22].OverrideCfg := 1, [2,23].TagName := 'SPARE', [2,23].Address := 23, [2,23].RawMin := 5529, [2,23].RawMax := 27648, [2,23].RealCfg := 1, [2,23].OverrideCfg := 1, [2,24].TagName := 'SPARE', [2,24].Address := 24, [2,24].RawMin := 5529, [2,24].RawMax := 27648, [2,24].RealCfg := 1, [2,24].OverrideCfg := 1, [2,25].TagName := 'SPARE', [2,25].Address := 25, [2,25].RawMin := 5529, [2,25].RawMax := 27648, [2,25].RealCfg := 1, [2,25].OverrideCfg := 1, [2,26].TagName := 'SPARE', [2,26].Address := 26, [2,26].RawMin := 5529, [2,26].RawMax := 27648, [2,26].RealCfg := 1,
        [2,26].OverrideCfg := 1, [2,27].TagName := 'SPARE', [2,27].Address := 27, [2,27].RawMin := 5529, [2,27].RawMax := 27648, [2,27].RealCfg := 1, [2,27].OverrideCfg := 1, [2,28].TagName := 'AI#1', [2,28].OutofRange := 1, [2,28].Address := 28, [2,28].RawMin := 6553, [2,28].RawMax := 32767, [2,28].RawLowLimit := 6225, [2,28].RawHighLimit := 33095, [2,28].FilterActual := 1.0, [2,28].ScaledMax := 100.0, [2,28].CurrentValue := -24.998093, [2,28].RangeMax := 100.0, [2,28].RangeMaxSave := 100.0, [2,28].RealCfg := 1, [2,28].EnableCfg := 1, [2,28].OverrideCfg := 1, [2,29].TagName := 'AI#2', [2,29].OutofRange := 1, [2,29].Address := 29, [2,29].RawMin := 6553, [2,29].RawMax := 32767, [2,29].RawLowLimit := 6225, [2,29].RawHighLimit := 33095, [2,29].FilterActual := 1.0, [2,29].ScaledMax := 100.0, [2,29].CurrentValue := -24.998093, [2,29].RangeMax := 100.0, [2,29].RangeMaxSave := 100.0, [2,29].RealCfg := 1, [2,29].EnableCfg := 1, [2,29].OverrideCfg := 1, [2,30].TagName := 'AI#3', [2,30].OutofRange := 1, [2,30].Address := 30, [2,30].RawMin := 6553, [2,30].RawMax := 32767, [2,30].RawValue := 49, [2,30].RawLowLimit := 6225, [2,30].RawHighLimit := 33095, [2,30].FilteredRaw := 49, [2,30].FilterActual := 1.0, [2,30].ScaledMax := 100.0, [2,30].CurrentValue := -24.811169, [2,30].RangeMax := 100.0, [2,30].RangeMaxSave := 100.0, [2,30].RealCfg := 1, [2,30].EnableCfg := 1, [2,30].OverrideCfg := 1, [2,31].TagName := 'AI#4', [2,31].OutofRange := 1, [2,31].Address := 31, [2,31].RawMin := 6553, [2,31].RawMax := 32767, [2,31].RawValue := 48,
        [2,31].RawLowLimit := 6225, [2,31].RawHighLimit := 33095, [2,31].FilteredRaw := 48, [2,31].FilterActual := 1.0, [2,31].ScaledMax := 100.0, [2,31].CurrentValue := -24.814985, [2,31].RangeMax := 100.0, [2,31].RangeMaxSave := 100.0, [2,31].RealCfg := 1, [2,31].EnableCfg := 1, [2,31].OverrideCfg := 1, [2,40].TagName := 'FI003', [2,40].Address := 40, [2,40].RawMin := 5529, [2,40].RawMax := 27648, [2,40].RawLowLimit := 5253, [2,40].RawHighLimit := 27924, [2,40].FilterActual := 1.0, [2,40].ScaledMax := 44.0, [2,40].RangeMax := 44.0, [2,40].RangeMaxSave := 44.0, [2,40].EnableCfg := 1, [2,40].OverrideCfg := 1, [2,41].TagName := 'LV003', [2,41].Address := 41, [2,41].RawMin := 6553, [2,41].RawMax := 32767, [2,41].RawLowLimit := 6225, [2,41].RawHighLimit := 33095, [2,41].FilterActual := 1.0, [2,41].ScaledMax := 9999.0, [2,41].RangeMax := 9999.0, [2,41].RangeMaxSave := 9999.0, [2,41].EnableCfg := 1, [2,41].OverrideCfg := 1, [2,42].TagName := 'LV001', [2,42].Address := 42, [2,42].RawMin := 6553, [2,42].RawMax := 32767, [2,42].RawLowLimit := 6225, [2,42].RawHighLimit := 33095, [2,42].FilterActual := 1.0, [2,42].ScaledMax := 9999.0, [2,42].RangeMax := 9999.0, [2,42].RangeMaxSave := 9999.0, [2,42].EnableCfg := 1, [2,42].OverrideCfg := 1, [2,43].TagName := 'LV002', [2,43].Address := 43, [2,43].RawMin := 6553, [2,43].RawMax := 32767, [2,43].RawLowLimit := 6225, [2,43].RawHighLimit := 33095, [2,43].FilterActual := 1.0, [2,43].ScaledMax := 9999.0, [2,43].RangeMax := 9999.0, [2,43].RangeMaxSave := 9999.0, [2,43].EnableCfg := 1, [2,43].OverrideCfg := 1, [2,44].Address := 44,
        [2,44].RawMin := 6553, [2,44].RawMax := 32767, [2,44].RawLowLimit := 6225, [2,44].RawHighLimit := 33095, [2,44].FilterActual := 1.0, [2,44].ScaledMax := 99999.0, [2,44].RangeMax := 99999.0, [2,44].RangeMaxSave := 99999.0, [2,45].Address := 42, [2,45].RawMin := 6553, [2,45].RawMax := 32767, [2,45].RawLowLimit := 6225, [2,45].RawHighLimit := 33095, [2,45].FilterActual := 1.0, [2,45].ScaledMin := -1.0, [2,45].ScaledMax := 5.0, [2,45].RangeMin := -1.0, [2,45].RangeMax := 5.0, [2,45].RangeMinSave := -1.0, [2,45].RangeMaxSave := 5.0, [2,45].OverrideCfg := 1, [3,0].OutofRange := 1, [3,0].RawMin := 6553, [3,0].RawMax := 32767, [3,0].RawLowLimit := 6225, [3,0].RawHighLimit := 33095, [3,0].FilterActual := 1.0, [3,0].RealCfg := 1, [3,0].EnableCfg := 1, [3,0].OverrideCfg := 1, [3,1].TagName := 'PI002', [3,1].TagDisplayName := 'PI002', [3,1].OutofRange := 1, [3,1].Address := 1, [3,1].RawMin := 5529, [3,1].RawMax := 27648, [3,1].RawLowLimit := 5253, [3,1].RawHighLimit := 27924, [3,1].FilterUser := 50, [3,1].FilterActual := 0.5, [3,1].ScaledMax := 6.0, [3,1].CurrentValue := -0.06111238, [3,1].RangeMax := 6.0, [3,1].RangeMaxSave := 6.0, [3,1].RealCfg := 1, [3,1].EnableCfg := 1, [3,1].OverrideCfg := 1, [3,1].Desc := 'Retentate Pressure', [3,1].EGU := 'bar', [3,2].TagName := 'PI101', [3,2].TagDisplayName := 'PI101', [3,2].OutofRange := 1, [3,2].Address := 2, [3,2].RawMin := 5529, [3,2].RawMax := 27648, [3,2].RawLowLimit := 5253, [3,2].RawHighLimit := 27924, [3,2].FilterUser := 50, [3,2].FilterActual := 0.5, [3,2].ScaledMax := 6.0,
        [3,2].CurrentValue := -0.03822385, [3,2].RangeMax := 6.0, [3,2].RangeMaxSave := 6.0, [3,2].RealCfg := 1, [3,2].EnableCfg := 1, [3,2].OverrideCfg := 1, [3,2].Desc := 'Filtrate Pressure', [3,2].EGU := 'bar', [3,3].TagName := 'PI006', [3,3].TagDisplayName := 'PI006', [3,3].OutofRange := 1, [3,3].Address := 3, [3,3].RawMin := 5529, [3,3].RawMax := 27648, [3,3].RawLowLimit := 5253, [3,3].RawHighLimit := 27924, [3,3].FilterActual := 1.0, [3,3].ScaledMax := 5.0, [3,3].CurrentValue := 0.2228261, [3,3].RangeMax := 5.0, [3,3].RangeMaxSave := 5.0, [3,3].RealCfg := 1, [3,3].EnableCfg := 1, [3,3].OverrideCfg := 1, [3,3].Desc := 'Feed Pump Pressure', [3,3].EGU := 'bar', [3,4].TagName := 'PI401', [3,4].TagDisplayName := 'PI401', [3,4].OutofRange := 1, [3,4].Address := 4, [3,4].RawMin := 5529, [3,4].RawMax := 27648, [3,4].RawLowLimit := 5253, [3,4].RawHighLimit := 27924, [3,4].FilterActual := 1.0, [3,4].ScaledMax := 6.0, [3,4].CurrentValue := -0.03387503, [3,4].RangeMax := 6.0, [3,4].RangeMaxSave := 6.0, [3,4].RealCfg := 1, [3,4].EnableCfg := 1, [3,4].OverrideCfg := 1, [3,4].Desc := 'Transfer Pump Pressure', [3,4].EGU := 'bar', [3,5].TagName := 'PI06', [3,5].TagDisplayName := 'PI06', [3,5].OutofRange := 1, [3,5].Address := 5, [3,5].RawMin := 5529, [3,5].RawMax := 27648, [3,5].RawLowLimit := 5253, [3,5].RawHighLimit := 27924, [3,5].FilterActual := 1.0, [3,5].ScaledMax := 100.0, [3,5].CurrentValue := 1.033333, [3,5].RangeMax := 100.0, [3,5].RangeMaxSave := 100.0, [3,5].RealCfg := 1, [3,5].EnableCfg := 1, [3,5].OverrideCfg := 1,
        [3,6].TagName := 'FI001', [3,6].TagDisplayName := 'FI001', [3,6].OutofRange := 1, [3,6].Address := 6, [3,6].RawMin := 5529, [3,6].RawMax := 27648, [3,6].RawLowLimit := 5253, [3,6].RawHighLimit := 27924, [3,6].FilterActual := 1.0, [3,6].ScaledMax := 25.0, [3,6].RangeMax := 25.0, [3,6].RangeMaxSave := 25.0, [3,6].RealCfg := 1, [3,6].EnableCfg := 1, [3,6].OverrideCfg := 1, [3,6].Desc := 'Calculated Feed Flow', [3,6].EGU := 'lpm', [3,7].TagName := 'FI101', [3,7].TagDisplayName := 'FI101', [3,7].OutofRange := 1, [3,7].Address := 7, [3,7].RawMin := 5529, [3,7].RawMax := 27648, [3,7].RawLowLimit := 5253, [3,7].RawHighLimit := 27924, [3,7].FilterActual := 1.0, [3,7].ScaledMax := 15.0, [3,7].RangeMax := 15.0, [3,7].RangeMaxSave := 15.0, [3,7].RealCfg := 1, [3,7].EnableCfg := 1, [3,7].OverrideCfg := 1, [3,7].Desc := 'Filtrate Flow', [3,7].EGU := 'lpm', [3,8].TagName := 'FI601', [3,8].TagDisplayName := 'FI601', [3,8].OutofRange := 1, [3,8].Address := 8, [3,8].RawMin := 5529, [3,8].RawMax := 27648, [3,8].RawLowLimit := 5253, [3,8].RawHighLimit := 27924, [3,8].FilterActual := 1.0, [3,8].ScaledMax := 2000.0, [3,8].CurrentValue := -25.10109, [3,8].RangeMax := 2000.0, [3,8].RangeMaxSave := 2000.0, [3,8].RealCfg := 1, [3,8].EnableCfg := 1, [3,8].OverrideCfg := 1, [3,8].Desc := 'Integrity Air Flow', [3,8].EGU := 'mlpm', [3,9].TagName := 'FI401', [3,9].TagDisplayName := 'FI401', [3,9].OutofRange := 1, [3,9].Address := 9, [3,9].RawMin := 6553, [3,9].RawMax := 32767, [3,9].RawLowLimit := 6225, [3,9].RawHighLimit := 33095,
        [3,9].FilterActual := 1.0, [3,9].ScaledMax := 25.0, [3,9].RangeMax := 25.0, [3,9].RangeMaxSave := 25.0, [3,9].RealCfg := 1, [3,9].EnableCfg := 1, [3,9].OverrideCfg := 1, [3,9].Desc := 'Calculated Trans Pump Flow', [3,9].EGU := 'lpm', [3,10].TagName := 'TI001', [3,10].TagDisplayName := 'TI001', [3,10].Address := 10, [3,10].RawMin := 5529, [3,10].RawMax := 27648, [3,10].RawLowLimit := 5253, [3,10].RawHighLimit := 27924, [3,10].FilterActual := 1.0, [3,10].ScaledMax := 55.0, [3,10].CurrentValue := 20.567827, [3,10].RangeMax := 55.0, [3,10].RangeMaxSave := 55.0, [3,10].EnableCfg := 1, [3,10].OverrideCfg := 1, [3,10].Desc := 'Feed Bag Temperature', [3,10].EGU := 'degC', [3,11].TagName := 'TI009', [3,11].TagDisplayName := 'TI009', [3,11].OutofRange := 1, [3,11].Address := 11, [3,11].RawMin := 6553, [3,11].RawMax := 32767, [3,11].RawLowLimit := 6225, [3,11].RawHighLimit := 33095, [3,11].FilterActual := 1.0, [3,11].ScaledMax := 30.0, [3,11].CurrentValue := 25.7337, [3,11].RangeMax := 30.0, [3,11].RangeMaxSave := 30.0, [3,11].RealCfg := 1, [3,11].EnableCfg := 1, [3,11].OverrideCfg := 1, [3,11].Desc := 'Retentate temperature', [3,11].EGU := 'degC', [3,12].TagName := 'TI012', [3,12].TagDisplayName := 'TI101', [3,12].Address := 12, [3,12].RawMin := 5529, [3,12].RawMax := 27648, [3,12].RawLowLimit := 5253, [3,12].RawHighLimit := 27924, [3,12].FilterActual := 1.0, [3,12].ScaledMax := 30.0, [3,12].CurrentValue := 28.0231, [3,12].RangeMax := 30.0, [3,12].RangeMaxSave := 30.0, [3,12].EnableCfg := 1, [3,12].OverrideCfg := 1, [3,12].Desc := 'Filtrate Temperature', [3,12].EGU := 'degC', [3,13].TagName := 'TI04',
        [3,13].TagDisplayName := 'TI04', [3,13].OutofRange := 1, [3,13].Address := 13, [3,13].RawMin := 6553, [3,13].RawMax := 32767, [3,13].RawLowLimit := 6225, [3,13].RawHighLimit := 33095, [3,13].FilterActual := 1.0, [3,13].ScaledMax := 150.0, [3,13].CurrentValue := 21.08868, [3,13].RangeMax := 150.0, [3,13].RangeMaxSave := 150.0, [3,13].RealCfg := 1, [3,13].EnableCfg := 1, [3,13].OverrideCfg := 1, [3,14].TagName := 'LI001', [3,14].TagDisplayName := 'LI001', [3,14].Address := 14, [3,14].RawMin := 6553, [3,14].RawMax := 32767, [3,14].RawValue := 20635, [3,14].RawLowLimit := 6225, [3,14].RawHighLimit := 33095, [3,14].FilteredRaw := 20635, [3,14].FilterActual := 1.0, [3,14].ScaledMax := 999.99, [3,14].CurrentValue := -0.04, [3,14].RangeMax := 240.0, [3,14].RangeMaxSave := 240.0, [3,14].Desc := 'Feed Bag Volume', [3,14].EGU := 'l', [3,15].TagName := 'WI101', [3,15].TagDisplayName := 'WI101', [3,15].OutofRange := 1, [3,15].Address := 15, [3,15].RawMax := 99999, [3,15].RawValue := 3, [3,15].RawLowLimit := -1000, [3,15].RawHighLimit := 100999, [3,15].FilterActual := 1.0, [3,15].ScaledMax := 9999.9, [3,15].CurrentValue := 0.29999793, [3,15].RangeMax := 600.0, [3,15].RangeMaxSave := 600.0, [3,15].RealCfg := 1, [3,15].Desc := 'Filtrate Weight', [3,15].EGU := 'kg', [3,16].TagName := 'WI102', [3,16].TagDisplayName := 'WI102', [3,16].OutofRange := 1, [3,16].Address := 16, [3,16].RawMin := 6553, [3,16].RawMax := 32767, [3,16].RawLowLimit := 6225, [3,16].RawHighLimit := 33095, [3,16].FilterActual := 1.0, [3,16].ScaledMax := 1000.0, [3,16].CurrentValue := -249.98116, [3,16].RangeMax := 1000.0, [3,16].RangeMaxSave := 1000.0,
        [3,16].RealCfg := 1, [3,16].Desc := 'Customer Filtrate Weight', [3,16].EGU := 'kg', [3,17].TagName := 'WI001', [3,17].TagDisplayName := 'WI001', [3,17].OutofRange := 1, [3,17].Address := 17, [3,17].RawMax := 99999, [3,17].RawValue := -4, [3,17].RawLowLimit := -1000, [3,17].RawHighLimit := 100999, [3,17].FilterActual := 1.0, [3,17].ScaledMax := 999.99, [3,17].CurrentValue := -0.04, [3,17].RangeMax := 240.0, [3,17].RangeMaxSave := 240.0, [3,17].RealCfg := 1, [3,17].Desc := 'Feed Bag Weight', [3,17].EGU := 'kg', [3,18].TagName := 'AI101', [3,18].TagDisplayName := 'AI101', [3,18].Address := 18, [3,18].RawMin := 6553, [3,18].RawMax := 32767, [3,18].RawValue := 32767, [3,18].RawLowLimit := 6225, [3,18].RawHighLimit := 33095, [3,18].FilteredRaw := 32767, [3,18].FilterActual := 1.0, [3,18].ScaledMax := 100.0, [3,18].CurrentValue := 100.0, [3,18].RangeMax := 100.0, [3,18].RangeMaxSave := 100.0, [3,18].RealCfg := 1, [3,18].Desc := 'Filtrate Conductivity', [3,18].EGU := 'uS', [3,19].TagName := 'AI102', [3,19].TagDisplayName := 'AI102', [3,19].Address := 19, [3,19].RawMin := 6553, [3,19].RawMax := 32767, [3,19].RawValue := 6446, [3,19].RawLowLimit := 6225, [3,19].RawHighLimit := 33095, [3,19].FilteredRaw := 6446, [3,19].FilterActual := 1.0, [3,19].ScaledMax := 2.0, [3,19].CurrentValue := -0.008163577, [3,19].RangeMax := 2.0, [3,19].RangeMaxSave := 2.0, [3,19].RealCfg := 1, [3,19].Desc := 'Filtrate UV', [3,19].EGU := 'AU', [3,20].TagName := 'AI103', [3,20].TagDisplayName := 'AI103', [3,20].Address := 20, [3,20].RawMin := 6553, [3,20].RawMax := 32767, [3,20].RawValue := 6429, [3,20].RawLowLimit := 6225,
        [3,20].RawHighLimit := 33095, [3,20].FilteredRaw := 6429, [3,20].FilterActual := 1.0, [3,20].ScaledMax := 2.0, [3,20].CurrentValue := -0.009460594, [3,20].RangeMax := 2.0, [3,20].RangeMaxSave := 2.0, [3,20].RealCfg := 1, [3,20].Desc := 'Filtrate UV', [3,20].EGU := 'AU', [3,21].TagName := 'AI104', [3,21].TagDisplayName := 'AI104', [3,21].OutofRange := 1, [3,21].Address := 21, [3,21].RawMin := 6553, [3,21].RawMax := 32767, [3,21].RawLowLimit := 6225, [3,21].RawHighLimit := 33095, [3,21].FilterActual := 1.0, [3,21].ScaledMax := 14.0, [3,21].CurrentValue := -3.499733, [3,21].RangeMax := 14.0, [3,21].RangeMaxSave := 14.0, [3,21].RealCfg := 1, [3,21].Desc := 'Filtrate pH', [3,21].EGU := 'pH', [3,22].TagName := 'AI010', [3,22].TagDisplayName := 'AI014', [3,22].Address := 22, [3,22].RawMin := 5520, [3,22].RawMax := 27600, [3,22].RawValue := 6592, [3,22].RawLowLimit := 5244, [3,22].RawHighLimit := 27876, [3,22].FilteredRaw := 6592, [3,22].FilterActual := 1.0, [3,22].ScaledMax := 3.0, [3,22].CurrentValue := 0.1456522, [3,22].RangeMax := 3.0, [3,22].RangeMaxSave := 3.0, [3,22].Desc := 'Retentate pH', [3,22].EGU := 'AU', [3,23].TagName := 'AI01', [3,23].TagDisplayName := 'AI01', [3,23].OutofRange := 1, [3,23].Address := 23, [3,23].RawMin := 6553, [3,23].RawMax := 32767, [3,23].RawLowLimit := 6225, [3,23].RawHighLimit := 33095, [3,23].FilterActual := 1.0, [3,23].ScaledMax := 100.0, [3,23].CurrentValue := -24.99809, [3,23].RangeMax := 100.0, [3,23].RangeMaxSave := 100.0, [3,23].Desc := 'Customer Input 01', [3,24].TagName := 'AI02', [3,24].TagDisplayName := 'AI02', [3,24].OutofRange := 1, [3,24].Address := 24,
        [3,24].RawMin := 6553, [3,24].RawMax := 32767, [3,24].RawLowLimit := 6225, [3,24].RawHighLimit := 33095, [3,24].FilterActual := 1.0, [3,24].ScaledMax := 100.0, [3,24].CurrentValue := -24.99809, [3,24].RangeMax := 100.0, [3,24].RangeMaxSave := 100.0, [3,24].RealCfg := 1, [3,24].Desc := 'Customer Input 02', [3,25].TagName := 'AI03', [3,25].TagDisplayName := 'AI03', [3,25].OutofRange := 1, [3,25].Address := 25, [3,25].RawMin := 6553, [3,25].RawMax := 32767, [3,25].RawLowLimit := 6225, [3,25].RawHighLimit := 33095, [3,25].FilterActual := 1.0, [3,25].ScaledMax := 100.0, [3,25].CurrentValue := -24.99809, [3,25].RangeMax := 100.0, [3,25].RangeMaxSave := 100.0, [3,25].RealCfg := 1, [3,25].Desc := 'Customer Input 03', [3,26].TagName := 'TI05', [3,26].TagDisplayName := 'TI05', [3,26].OutofRange := 1, [3,26].Address := 26, [3,26].RawMin := 6553, [3,26].RawMax := 32767, [3,26].RawValue := 8, [3,26].RawLowLimit := 6225, [3,26].RawHighLimit := 33095, [3,26].FilteredRaw := 8, [3,26].FilterActual := 1.0, [3,26].CurrentValue := 63.88032, [3,26].RealCfg := 1, [3,27].TagName := 'TI06', [3,27].TagDisplayName := 'TI06', [3,27].Address := 27, [3,27].RawMin := 6553, [3,27].RawMax := 32767, [3,27].RawValue := 9728, [3,27].RawLowLimit := 6225, [3,27].RawHighLimit := 33095, [3,27].FilteredRaw := 9728, [3,27].FilterActual := 1.0, [3,27].ScaledMax := 150.0, [3,27].CurrentValue := 20.94448, [3,27].RangeMax := 150.0, [3,27].RangeMaxSave := 150.0, [3,27].RealCfg := 1, [3,28].TagName := 'PCV001', [3,28].TagDisplayName := 'PCV001', [3,28].OutofRange := 1, [3,28].Address := 28, [3,28].RawMin := 6553, [3,28].RawMax := 32767,
        [3,28].RawLowLimit := 6225, [3,28].RawHighLimit := 33095, [3,28].FilterActual := 1.0, [3,28].ScaledMax := 100.0, [3,28].CurrentValue := -1.048729, [3,28].RangeMax := 100.0, [3,28].RangeMaxSave := 100.0, [3,28].RealCfg := 1, [3,28].EnableCfg := 1, [3,28].OverrideCfg := 1, [3,28].Desc := 'Retentate Pressure Valve', [3,28].EGU := '%', [3,29].TagName := 'PCV101', [3,29].TagDisplayName := 'PCV101', [3,29].OutofRange := 1, [3,29].Address := 29, [3,29].RawMin := 6553, [3,29].RawMax := 32767, [3,29].RawLowLimit := 6225, [3,29].RawHighLimit := 33095, [3,29].FilterActual := 1.0, [3,29].ScaledMax := 100.0, [3,29].CurrentValue := 100.96327, [3,29].RangeMax := 100.0, [3,29].RangeMaxSave := 100.0, [3,29].RealCfg := 1, [3,29].EnableCfg := 1, [3,29].OverrideCfg := 1, [3,29].Desc := 'Filtrate Pressure Valve', [3,29].EGU := '%', [3,30].TagName := 'MIX001', [3,30].TagDisplayName := 'MIX001', [3,30].OutofRange := 1, [3,30].Address := 30, [3,30].RawMin := 6553, [3,30].RawMax := 32767, [3,30].RawLowLimit := 6225, [3,30].RawHighLimit := 33095, [3,30].FilterActual := 1.0, [3,30].ScaledMax := 100.0, [3,30].CurrentValue := 0.024414062, [3,30].RangeMax := 100.0, [3,30].RangeMaxSave := 100.0, [3,30].RealCfg := 1, [3,30].EnableCfg := 1, [3,30].OverrideCfg := 1, [3,30].Desc := 'Mixer Speed', [3,30].EGU := '%', [3,31].TagName := 'AP31', [3,31].TagDisplayName := 'AP31', [3,31].OutofRange := 1, [3,31].Address := 31, [3,31].RawMin := 6553, [3,31].RawMax := 32767, [3,31].RawLowLimit := 6225, [3,31].RawHighLimit := 33095, [3,31].FilterActual := 1.0, [3,31].ScaledMax := 100.0, [3,31].CurrentValue := 9.026997, [3,31].RangeMax := 100.0,
        [3,31].RangeMaxSave := 100.0, [3,31].RealCfg := 1, [3,31].EnableCfg := 1, [3,31].OverrideCfg := 1, [3,32].TagName := 'DP', [3,32].TagDisplayName := 'DP', [3,32].Address := 32, [3,32].FilterActual := 1.0, [3,32].ScaledMax := 6.0, [3,32].CurrentValue := 0.045777064, [3,32].RangeMax := 6.0, [3,32].RangeMaxSave := 6.0, [3,32].Desc := 'Differential Pressure', [3,32].EGU := 'bar', [3,33].TagName := 'TMP', [3,33].TagDisplayName := 'TMP', [3,33].Address := 33, [3,33].FilterActual := 1.0, [3,33].ScaledMax := 6.0, [3,33].CurrentValue := 3.7252903e-09, [3,33].RangeMax := 6.0, [3,33].RangeMaxSave := 6.0, [3,33].Desc := 'Trans-Membrane Pressure', [3,33].EGU := 'bar', [3,34].TagName := 'PD03', [3,34].TagDisplayName := 'PD03', [3,34].Address := 34, [3,34].RawValue := 6248, [3,34].FilteredRaw := 6248, [3,34].FilterActual := 1.0, [3,34].ScaledMax := 100.0, [3,34].CurrentValue := 0.06248569, [3,34].RangeMax := 100.0, [3,34].RangeMaxSave := 100.0, [3,35].TagName := 'FI04', [3,35].TagDisplayName := 'FI04', [3,35].Address := 35, [3,35].RawMin := 6553, [3,35].RawMax := 32767, [3,35].RawLowLimit := 6225, [3,35].RawHighLimit := 33095, [3,35].FilterActual := 1.0, [3,35].ScaledMax := 100.0, [3,35].CurrentValue := 222.0, [3,35].RangeMax := 100.0, [3,35].RangeMaxSave := 100.0, [3,36].TagName := 'LV', [3,36].Address := 36, [3,36].RawMin := 6553, [3,36].RawMax := 32767, [3,36].RawLowLimit := 6225, [3,36].RawHighLimit := 33095, [3,36].FilterActual := 1.0, [3,36].ScaledMax := 1000.0, [3,36].RangeMax := 1000.0, [3,36].RangeMaxSave := 1000.0, [3,36].EGU := 'cmhr', [3,37].TagName := 'PI001', [3,37].TagDisplayName := 'PI001', [3,37].Address := 37,
        [3,37].RawMin := 6553, [3,37].RawMax := 32767, [3,37].RawValue := 6486, [3,37].RawLowLimit := 6225, [3,37].RawHighLimit := 33095, [3,37].FilterUser := 50, [3,37].FilteredRaw := 6486, [3,37].FilterActual := 0.5, [3,37].ScaledMax := 6.0, [3,37].CurrentValue := -0.015335317, [3,37].RangeMax := 6.0, [3,37].RangeMaxSave := 6.0, [3,37].RealCfg := 1, [3,37].Desc := 'Feed Pressure', [3,37].EGU := 'bar', [3,38].TagName := 'NWP', [3,38].TagDisplayName := 'NWP', [3,38].FilterActual := 1.0, [3,38].ScaledMax := 1000.0, [3,38].RangeMax := 1000.0, [3,38].RangeMaxSave := 1000.0, [3,38].EGU := 'lm2h/', [3,39].TagName := 'PERM', [3,39].TagDisplayName := 'PERM', [3,39].FilterActual := 1.0, [3,39].ScaledMax := 1000.0, [3,39].RangeMax := 1000.0, [3,39].RangeMaxSave := 1000.0, [3,39].EGU := 'lm2/', [3,40].Address := 40, [3,40].RawMin := 5529, [3,40].RawMax := 27648, [3,40].RawLowLimit := 5253, [3,40].RawHighLimit := 27924, [3,40].FilterActual := 1.0, [3,40].CurrentValue := 48.590927, [3,40].EnableCfg := 1, [3,40].OverrideCfg := 1, [3,41].Address := 41, [3,41].RawMin := 6553, [3,41].RawMax := 32767, [3,41].RawLowLimit := 6225, [3,41].RawHighLimit := 33095, [3,41].FilterActual := 1.0, [3,41].CurrentValue := 5830.911, [3,41].EnableCfg := 1, [3,41].OverrideCfg := 1, [3,42].Address := 42, [3,42].RawMin := 6553, [3,42].RawMax := 32767, [3,42].RawLowLimit := 6225, [3,42].RawHighLimit := 33095, [3,42].FilterActual := 1.0, [3,42].CurrentValue := 2468.1392, [3,42].EnableCfg := 1, [3,42].OverrideCfg := 1, [3,43].Address := 43, [3,43].RawMin := 6553, [3,43].RawMax := 32767, [3,43].RawLowLimit := 6225,
        [3,43].RawHighLimit := 33095, [3,43].FilterActual := 1.0, [3,43].CurrentValue := 3362.772, [3,43].EnableCfg := 1, [3,43].OverrideCfg := 1, [4,0].TagName := 'PCV032', [4,0].OutofRange := 1, [4,0].FilterActual := 1.0, [4,0].ScaledMax := 100.0, [4,0].RangeMax := 100.0, [4,0].RangeMaxSave := 100.0, [4,0].RealCfg := 1, [4,0].EnableCfg := 1, [4,0].OverrideCfg := 1, [4,1].TagName := 'AI201B', [4,1].OutofRange := 1, [4,1].Address := 1, [4,1].RawMin := 5529, [4,1].RawMax := 27648, [4,1].RawLowLimit := 5253, [4,1].RawHighLimit := 27924, [4,1].FilterActual := 1.0, [4,1].ScaledMax := 50.0, [4,1].CurrentValue := -12.498303, [4,1].RangeMax := 50.0, [4,1].RangeMaxSave := 50.0, [4,1].RealCfg := 1, [4,1].EnableCfg := 1, [4,1].OverrideCfg := 1, [4,2].TagName := 'AI201A', [4,2].OutofRange := 1, [4,2].Address := 2, [4,2].RawMin := 5529, [4,2].RawMax := 27648, [4,2].RawLowLimit := 5253, [4,2].RawHighLimit := 27924, [4,2].FilterActual := 1.0, [4,2].ScaledMax := 100.0, [4,2].CurrentValue := -24.996607, [4,2].RangeMax := 100.0, [4,2].RangeMaxSave := 100.0, [4,2].RealCfg := 1, [4,2].EnableCfg := 1, [4,2].OverrideCfg := 1, [4,3].TagName := 'AI202', [4,3].OutofRange := 1, [4,3].Address := 3, [4,3].RawMin := 5529, [4,3].RawMax := 27648, [4,3].RawLowLimit := 5253, [4,3].RawHighLimit := 27924, [4,3].FilterActual := 1.0, [4,3].ScaledMax := 14.0, [4,3].CurrentValue := -3.499525, [4,3].RangeMax := 14.0, [4,3].RangeMaxSave := 14.0, [4,3].RealCfg := 1, [4,3].EnableCfg := 1, [4,3].OverrideCfg := 1, [4,4].TagName := 'TI201',
        [4,4].OutofRange := 1, [4,4].Address := 4, [4,4].RawMin := 5529, [4,4].RawMax := 27648, [4,4].RawLowLimit := 5253, [4,4].RawHighLimit := 27924, [4,4].FilterActual := 1.0, [4,4].ScaledMax := 100.0, [4,4].CurrentValue := -24.996607, [4,4].RangeMax := 100.0, [4,4].RangeMaxSave := 100.0, [4,4].RealCfg := 1, [4,4].EnableCfg := 1, [4,4].OverrideCfg := 1, [4,5].TagName := 'AI203', [4,5].OutofRange := 1, [4,5].Address := 5, [4,5].RawMin := 5529, [4,5].RawMax := 27648, [4,5].RawLowLimit := 5253, [4,5].RawHighLimit := 27924, [4,5].FilterActual := 1.0, [4,5].ScaledMax := 3.0, [4,5].CurrentValue := -0.7498982, [4,5].RangeMax := 3.0, [4,5].RangeMaxSave := 3.0, [4,5].RealCfg := 1, [4,5].EnableCfg := 1, [4,5].OverrideCfg := 1, [4,6].TagName := 'AI204', [4,6].OutofRange := 1, [4,6].Address := 6, [4,6].RawMin := 5529, [4,6].RawMax := 27648, [4,6].RawLowLimit := 5253, [4,6].RawHighLimit := 27924, [4,6].FilterActual := 1.0, [4,6].ScaledMax := 2.0, [4,6].CurrentValue := -0.49993217, [4,6].RangeMax := 2.0, [4,6].RangeMaxSave := 2.0, [4,6].RealCfg := 1, [4,6].EnableCfg := 1, [4,6].OverrideCfg := 1, [4,7].TagName := 'AI102', [4,7].OutofRange := 1, [4,7].Address := 7, [4,7].RawMin := 5529, [4,7].RawMax := 27648, [4,7].RawLowLimit := 5253, [4,7].RawHighLimit := 27924, [4,7].FilterActual := 1.0, [4,7].ScaledMax := 100.0, [4,7].CurrentValue := -24.996607, [4,7].RangeMax := 100.0, [4,7].RangeMaxSave := 100.0, [4,7].RealCfg := 1, [4,7].EnableCfg := 1, [4,7].OverrideCfg := 1, [4,8].TagName := 'AI103',
        [4,8].OutofRange := 1, [4,8].Address := 8, [4,8].RawMin := 5529, [4,8].RawMax := 27648, [4,8].RawLowLimit := 5253, [4,8].RawHighLimit := 27924, [4,8].FilterActual := 1.0, [4,8].ScaledMax := 14.0, [4,8].CurrentValue := -3.499525, [4,8].RangeMax := 14.0, [4,8].RangeMaxSave := 14.0, [4,8].RealCfg := 1, [4,8].EnableCfg := 1, [4,8].OverrideCfg := 1, [4,9].TagName := 'PI003', [4,9].OutofRange := 1, [4,9].Address := 9, [4,9].RawMin := 6553, [4,9].RawMax := 32767, [4,9].RawLowLimit := 6225, [4,9].RawHighLimit := 33095, [4,9].FilterActual := 1.0, [4,9].ScaledMax := 6.0, [4,9].CurrentValue := -1.4998856, [4,9].RangeMax := 6.0, [4,9].RangeMaxSave := 6.0, [4,9].RealCfg := 1, [4,9].EnableCfg := 1, [4,9].OverrideCfg := 1, [4,10].TagName := 'FI001', [4,10].OutofRange := 1, [4,10].Address := 10, [4,10].RawMin := 5529, [4,10].RawMax := 27648, [4,10].RawLowLimit := 5253, [4,10].RawHighLimit := 27924, [4,10].FilterActual := 1.0, [4,10].ScaledMax := 22.0, [4,10].RangeMax := 22.0, [4,10].RangeMaxSave := 22.0, [4,10].EnableCfg := 1, [4,10].OverrideCfg := 1, [4,11].TagName := 'PI001', [4,11].OutofRange := 1, [4,11].Address := 11, [4,11].RawMin := 6553, [4,11].RawMax := 32767, [4,11].RawLowLimit := 6225, [4,11].RawHighLimit := 33095, [4,11].FilterActual := 1.0, [4,11].ScaledMax := 6.0, [4,11].CurrentValue := -1.4998856, [4,11].RangeMax := 6.0, [4,11].RangeMaxSave := 6.0, [4,11].RealCfg := 1, [4,11].EnableCfg := 1, [4,11].OverrideCfg := 1, [4,12].TagName := 'FI002', [4,12].OutofRange := 1, [4,12].Address := 12,
        [4,12].RawMin := 5529, [4,12].RawMax := 27648, [4,12].RawLowLimit := 5253, [4,12].RawHighLimit := 27924, [4,12].FilterActual := 1.0, [4,12].ScaledMax := 22.0, [4,12].RangeMax := 22.0, [4,12].RangeMaxSave := 22.0, [4,12].EnableCfg := 1, [4,12].OverrideCfg := 1, [4,13].TagName := 'PI002', [4,13].OutofRange := 1, [4,13].Address := 13, [4,13].RawMin := 6553, [4,13].RawMax := 32767, [4,13].RawLowLimit := 6225, [4,13].RawHighLimit := 33095, [4,13].FilterActual := 1.0, [4,13].ScaledMax := 6.0, [4,13].CurrentValue := -1.4998856, [4,13].RangeMax := 6.0, [4,13].RangeMaxSave := 6.0, [4,13].RealCfg := 1, [4,13].EnableCfg := 1, [4,13].OverrideCfg := 1, [4,14].OutofRange := 1, [4,14].Address := 14, [4,14].RawMin := 5529, [4,14].RawMax := 27648, [4,14].RawLowLimit := 5253, [4,14].RawHighLimit := 27924, [4,14].FilterActual := 1.0, [4,14].ScaledMax := 14.0, [4,14].RangeMax := 14.0, [4,14].RangeMaxSave := 14.0, [4,14].RealCfg := 1, [4,14].OverrideCfg := 1, [4,15].OutofRange := 1, [4,15].Address := 15, [4,15].RawMin := 5529, [4,15].RawMax := 27648, [4,15].RawLowLimit := 5253, [4,15].RawHighLimit := 27924, [4,15].FilterActual := 1.0, [4,15].ScaledMax := 2.0, [4,15].CurrentValue := -0.49993217, [4,15].RangeMax := 2.0, [4,15].RangeMaxSave := 2.0, [4,15].RealCfg := 1, [4,15].OverrideCfg := 1, [4,16].OutofRange := 1, [4,16].Address := 16, [4,16].RawMin := 5529, [4,16].RawMax := 27648, [4,16].RawLowLimit := 5253, [4,16].RawHighLimit := 27924, [4,16].FilterActual := 1.0, [4,16].ScaledMax := 2.0, [4,16].CurrentValue := -0.49993217, [4,16].RangeMax := 2.0,
        [4,16].RangeMaxSave := 2.0, [4,16].RealCfg := 1, [4,16].OverrideCfg := 1, [4,17].OutofRange := 1, [4,17].Address := 17, [4,17].RawMin := 5529, [4,17].RawMax := 27648, [4,17].RawLowLimit := 5253, [4,17].RawHighLimit := 27924, [4,17].FilterActual := 1.0, [4,17].ScaledMin := -1.0, [4,17].ScaledMax := 5.0, [4,17].CurrentValue := -2.4997964, [4,17].RangeMin := -1.0, [4,17].RangeMax := 5.0, [4,17].RangeMinSave := -1.0, [4,17].RangeMaxSave := 5.0, [4,17].RealCfg := 1, [4,17].OverrideCfg := 1, [4,18].OutofRange := 1, [4,18].Address := 18, [4,18].RawMin := 5529, [4,18].RawMax := 27648, [4,18].RawLowLimit := 5253, [4,18].RawHighLimit := 27924, [4,18].FilterActual := 1.0, [4,18].ScaledMin := -1.0, [4,18].ScaledMax := 5.0, [4,18].CurrentValue := -2.4997964, [4,18].RangeMin := -1.0, [4,18].RangeMax := 5.0, [4,18].RangeMinSave := -1.0, [4,18].RangeMaxSave := 5.0, [4,18].RealCfg := 1, [4,18].OverrideCfg := 1, [4,19].OutofRange := 1, [4,19].Address := 19, [4,19].RawMin := 5529, [4,19].RawMax := 27648, [4,19].RawLowLimit := 5253, [4,19].RawHighLimit := 27924, [4,19].FilterActual := 1.0, [4,19].ScaledMin := -1.0, [4,19].ScaledMax := 5.0, [4,19].CurrentValue := -2.4997964, [4,19].RangeMin := -1.0, [4,19].RangeMax := 5.0, [4,19].RangeMinSave := -1.0, [4,19].RangeMaxSave := 5.0, [4,19].RealCfg := 1, [4,19].OverrideCfg := 1, [4,20].OutofRange := 1, [4,20].Address := 20, [4,20].RawMin := 5529, [4,20].RawMax := 27648, [4,20].RawLowLimit := 5253, [4,20].RawHighLimit := 27924, [4,20].FilterActual := 1.0, [4,20].ScaledMax := 100.0, [4,20].CurrentValue := -24.996607,
        [4,20].RangeMax := 100.0, [4,20].RangeMaxSave := 100.0, [4,20].RealCfg := 1, [4,20].OverrideCfg := 1, [4,21].OutofRange := 1, [4,21].Address := 21, [4,21].RawMin := 5529, [4,21].RawMax := 27648, [4,21].RawLowLimit := 5253, [4,21].RawHighLimit := 27924, [4,21].FilterActual := 1.0, [4,21].ScaledMax := 100.0, [4,21].CurrentValue := -24.996607, [4,21].RangeMax := 100.0, [4,21].RangeMaxSave := 100.0, [4,21].RealCfg := 1, [4,21].OverrideCfg := 1, [4,22].TagName := 'SPARE', [4,22].Address := 22, [4,22].RawMin := 5529, [4,22].RawMax := 27648, [4,22].RealCfg := 1, [4,22].OverrideCfg := 1, [4,23].TagName := 'SPARE', [4,23].Address := 23, [4,23].RawMin := 5529, [4,23].RawMax := 27648, [4,23].RealCfg := 1, [4,23].OverrideCfg := 1, [4,24].TagName := 'SPARE', [4,24].Address := 24, [4,24].RawMin := 5529, [4,24].RawMax := 27648, [4,24].RealCfg := 1, [4,24].OverrideCfg := 1, [4,25].TagName := 'SPARE', [4,25].Address := 25, [4,25].RawMin := 5529, [4,25].RawMax := 27648, [4,25].RealCfg := 1, [4,25].OverrideCfg := 1, [4,26].TagName := 'SPARE', [4,26].Address := 26, [4,26].RawMin := 5529, [4,26].RawMax := 27648, [4,26].RealCfg := 1, [4,26].OverrideCfg := 1, [4,27].TagName := 'SPARE', [4,27].Address := 27, [4,27].RawMin := 5529, [4,27].RawMax := 27648, [4,27].RealCfg := 1, [4,27].OverrideCfg := 1, [4,28].TagName := 'AI#1', [4,28].Address := 28, [4,28].RawMin := 6553, [4,28].RawMax := 32767, [4,28].RawValue := 12544, [4,28].RawLowLimit := 6225, [4,28].RawHighLimit := 33095,
        [4,28].FilteredRaw := 12544, [4,28].FilterActual := 1.0, [4,28].ScaledMax := 100.0, [4,28].CurrentValue := 22.8542, [4,28].RangeMax := 100.0, [4,28].RangeMaxSave := 100.0, [4,28].RealCfg := 1, [4,28].EnableCfg := 1, [4,28].OverrideCfg := 1, [4,29].TagName := 'AI#2', [4,29].Address := 29, [4,29].RawMin := 6553, [4,29].RawMax := 32767, [4,29].RawValue := 12288, [4,29].RawLowLimit := 6225, [4,29].RawHighLimit := 33095, [4,29].FilteredRaw := 12288, [4,29].FilterActual := 1.0, [4,29].ScaledMax := 100.0, [4,29].CurrentValue := 21.877623, [4,29].RangeMax := 100.0, [4,29].RangeMaxSave := 100.0, [4,29].RealCfg := 1, [4,29].EnableCfg := 1, [4,29].OverrideCfg := 1, [4,30].TagName := 'AI#3', [4,30].Address := 30, [4,30].RawMin := 6553, [4,30].RawMax := 32767, [4,30].RawValue := 12288, [4,30].RawLowLimit := 6225, [4,30].RawHighLimit := 33095, [4,30].FilteredRaw := 12288, [4,30].FilterActual := 1.0, [4,30].ScaledMax := 100.0, [4,30].CurrentValue := 21.877623, [4,30].RangeMax := 100.0, [4,30].RangeMaxSave := 100.0, [4,30].RealCfg := 1, [4,30].EnableCfg := 1, [4,30].OverrideCfg := 1, [4,31].TagName := 'AI#4', [4,31].Address := 31, [4,31].RawMin := 6553, [4,31].RawMax := 32767, [4,31].RawValue := 12288, [4,31].RawLowLimit := 6225, [4,31].RawHighLimit := 33095, [4,31].FilteredRaw := 12288, [4,31].FilterActual := 1.0, [4,31].ScaledMax := 100.0, [4,31].CurrentValue := 21.877623, [4,31].RangeMax := 100.0, [4,31].RangeMaxSave := 100.0, [4,31].RealCfg := 1, [4,31].EnableCfg := 1, [4,31].OverrideCfg := 1, [4,40].TagName := 'FI003', [4,40].Address := 40, [4,40].RawMin := 5529,
        [4,40].RawMax := 27648, [4,40].RawLowLimit := 5253, [4,40].RawHighLimit := 27924, [4,40].FilterActual := 1.0, [4,40].ScaledMax := 44.0, [4,40].RangeMax := 44.0, [4,40].RangeMaxSave := 44.0, [4,40].EnableCfg := 1, [4,40].OverrideCfg := 1, [4,41].TagName := 'LV003', [4,41].Address := 41, [4,41].RawMin := 6553, [4,41].RawMax := 32767, [4,41].RawLowLimit := 6225, [4,41].RawHighLimit := 33095, [4,41].FilterActual := 1.0, [4,41].ScaledMax := 9999.0, [4,41].RangeMax := 9999.0, [4,41].RangeMaxSave := 9999.0, [4,41].EnableCfg := 1, [4,41].OverrideCfg := 1, [4,42].TagName := 'LV001', [4,42].Address := 42, [4,42].RawMin := 6553, [4,42].RawMax := 32767, [4,42].RawLowLimit := 6225, [4,42].RawHighLimit := 33095, [4,42].FilterActual := 1.0, [4,42].ScaledMax := 9999.0, [4,42].RangeMax := 9999.0, [4,42].RangeMaxSave := 9999.0, [4,42].EnableCfg := 1, [4,42].OverrideCfg := 1, [4,43].TagName := 'LV002', [4,43].Address := 43, [4,43].RawMin := 6553, [4,43].RawMax := 32767, [4,43].RawLowLimit := 6225, [4,43].RawHighLimit := 33095, [4,43].FilterActual := 1.0, [4,43].ScaledMax := 9999.0, [4,43].RangeMax := 9999.0, [4,43].RangeMaxSave := 9999.0, [4,43].EnableCfg := 1, [4,43].OverrideCfg := 1, [4,44].Address := 44, [4,44].RawMin := 6553, [4,44].RawMax := 32767, [4,44].RawLowLimit := 6225, [4,44].RawHighLimit := 33095, [4,44].FilterActual := 1.0, [4,44].ScaledMax := 99999.0, [4,44].RangeMax := 99999.0, [4,44].RangeMaxSave := 99999.0, [4,45].Address := 42, [4,45].RawMin := 6553, [4,45].RawMax := 32767, [4,45].RawLowLimit := 6225, [4,45].RawHighLimit := 33095, [4,45].FilterActual := 1.0,
        [4,45].ScaledMin := -1.0, [4,45].ScaledMax := 5.0, [4,45].RangeMin := -1.0, [4,45].RangeMax := 5.0, [4,45].RangeMinSave := -1.0, [4,45].RangeMaxSave := 5.0, [4,45].OverrideCfg := 1, [5,0].TagName := 'PCV032', [5,0].OutofRange := 1, [5,0].RawMin := 6553, [5,0].RawMax := 32767, [5,0].RawLowLimit := 6225, [5,0].RawHighLimit := 33095, [5,0].FilterActual := 1.0, [5,0].ScaledMin := -1.0, [5,0].ScaledMax := 5.0, [5,0].CurrentValue := -2.4998856, [5,0].RangeMin := -1.0, [5,0].RangeMax := 5.0, [5,0].RangeMinSave := -1.0, [5,0].RangeMaxSave := 5.0, [5,0].RealCfg := 1, [5,0].EnableCfg := 1, [5,0].OverrideCfg := 1, [5,1].TagName := 'AI201B', [5,1].OutofRange := 1, [5,1].Address := 1, [5,1].RawMin := 5529, [5,1].RawMax := 27648, [5,1].RawLowLimit := 5253, [5,1].RawHighLimit := 27924, [5,1].FilterActual := 1.0, [5,1].ScaledMax := 25.0, [5,1].CurrentValue := -6.249152, [5,1].RangeMax := 25.0, [5,1].RangeMaxSave := 25.0, [5,1].RealCfg := 1, [5,1].EnableCfg := 1, [5,1].OverrideCfg := 1, [5,2].TagName := 'AI201A', [5,2].OutofRange := 1, [5,2].Address := 2, [5,2].RawMin := 5529, [5,2].RawMax := 27648, [5,2].RawLowLimit := 5253, [5,2].RawHighLimit := 27924, [5,2].FilterActual := 1.0, [5,2].ScaledMin := -1.0, [5,2].ScaledMax := 5.0, [5,2].CurrentValue := -2.4997966, [5,2].RangeMin := -1.0, [5,2].RangeMax := 5.0, [5,2].RangeMinSave := -1.0, [5,2].RangeMaxSave := 5.0, [5,2].RealCfg := 1, [5,2].EnableCfg := 1, [5,2].OverrideCfg := 1, [5,3].TagName := 'AI202', [5,3].OutofRange := 1, [5,3].Address := 3,
        [5,3].RawMin := 5529, [5,3].RawMax := 27648, [5,3].RawLowLimit := 5253, [5,3].RawHighLimit := 27924, [5,3].FilterActual := 1.0, [5,3].ScaledMax := 25.0, [5,3].CurrentValue := -6.249152, [5,3].RangeMax := 25.0, [5,3].RangeMaxSave := 25.0, [5,3].RealCfg := 1, [5,3].EnableCfg := 1, [5,3].OverrideCfg := 1, [5,4].TagName := 'TI201', [5,4].OutofRange := 1, [5,4].Address := 4, [5,4].RawMin := 5529, [5,4].RawMax := 27648, [5,4].RawLowLimit := 5253, [5,4].RawHighLimit := 27924, [5,4].FilterActual := 1.0, [5,4].ScaledMax := 150.0, [5,4].CurrentValue := -37.49491, [5,4].RangeMax := 150.0, [5,4].RangeMaxSave := 150.0, [5,4].RealCfg := 1, [5,4].EnableCfg := 1, [5,4].OverrideCfg := 1, [5,5].TagName := 'AI203', [5,5].OutofRange := 1, [5,5].Address := 5, [5,5].RawMin := 5529, [5,5].RawMax := 27648, [5,5].RawLowLimit := 5253, [5,5].RawHighLimit := 27924, [5,5].FilterActual := 1.0, [5,5].ScaledMax := 150.0, [5,5].CurrentValue := -37.49491, [5,5].RangeMax := 150.0, [5,5].RangeMaxSave := 150.0, [5,5].RealCfg := 1, [5,5].EnableCfg := 1, [5,5].OverrideCfg := 1, [5,6].TagName := 'AI204', [5,6].OutofRange := 1, [5,6].Address := 6, [5,6].RawMin := 5529, [5,6].RawMax := 27648, [5,6].RawLowLimit := 5253, [5,6].RawHighLimit := 27924, [5,6].FilterActual := 1.0, [5,6].ScaledMin := -1.0, [5,6].ScaledMax := 5.0, [5,6].CurrentValue := -2.4997966, [5,6].RangeMin := -1.0, [5,6].RangeMax := 5.0, [5,6].RangeMinSave := -1.0, [5,6].RangeMaxSave := 5.0, [5,6].RealCfg := 1, [5,6].EnableCfg := 1, [5,6].OverrideCfg := 1,
        [5,7].TagName := 'AI102', [5,7].OutofRange := 1, [5,7].Address := 7, [5,7].RawMin := 5529, [5,7].RawMax := 27648, [5,7].RawLowLimit := 5253, [5,7].RawHighLimit := 27924, [5,7].FilterActual := 1.0, [5,7].ScaledMin := -1.0, [5,7].ScaledMax := 5.0, [5,7].CurrentValue := -2.4997966, [5,7].RangeMin := -1.0, [5,7].RangeMax := 5.0, [5,7].RangeMinSave := -1.0, [5,7].RangeMaxSave := 5.0, [5,7].RealCfg := 1, [5,7].EnableCfg := 1, [5,7].OverrideCfg := 1, [5,8].TagName := 'AI103', [5,8].OutofRange := 1, [5,8].Address := 8, [5,8].RawMin := 5529, [5,8].RawMax := 27648, [5,8].RawLowLimit := 5253, [5,8].RawHighLimit := 27924, [5,8].FilterActual := 1.0, [5,8].ScaledMax := 200.0, [5,8].CurrentValue := -49.993217, [5,8].RangeMax := 200.0, [5,8].RangeMaxSave := 200.0, [5,8].RealCfg := 1, [5,8].EnableCfg := 1, [5,8].OverrideCfg := 1, [5,9].TagName := 'PI003', [5,9].OutofRange := 1, [5,9].Address := 9, [5,9].RawMin := 6553, [5,9].RawMax := 32767, [5,9].RawLowLimit := 6225, [5,9].RawHighLimit := 33095, [5,9].FilterActual := 1.0, [5,9].ScaledMax := 14.0, [5,9].CurrentValue := -3.499733, [5,9].RangeMax := 14.0, [5,9].RangeMaxSave := 14.0, [5,9].RealCfg := 1, [5,9].EnableCfg := 1, [5,9].OverrideCfg := 1, [5,10].TagName := 'FI001', [5,10].Address := 10, [5,10].RawMin := 5529, [5,10].RawMax := 27648, [5,10].RawLowLimit := 5253, [5,10].RawHighLimit := 27924, [5,10].FilterActual := 1.0, [5,10].EnableCfg := 1, [5,10].OverrideCfg := 1, [5,11].TagName := 'PI001', [5,11].OutofRange := 1, [5,11].Address := 11,
        [5,11].RawMin := 6553, [5,11].RawMax := 32767, [5,11].RawLowLimit := 6225, [5,11].RawHighLimit := 33095, [5,11].FilterActual := 1.0, [5,11].ScaledMax := 200.0, [5,11].CurrentValue := -49.996185, [5,11].RangeMax := 200.0, [5,11].RangeMaxSave := 200.0, [5,11].RealCfg := 1, [5,11].EnableCfg := 1, [5,11].OverrideCfg := 1, [5,12].TagName := 'FI002', [5,12].Address := 12, [5,12].RawMin := 5529, [5,12].RawMax := 27648, [5,12].RawLowLimit := 5253, [5,12].RawHighLimit := 27924, [5,12].FilterActual := 1.0, [5,12].ScaledMax := 50.0, [5,12].RangeMax := 50.0, [5,12].RangeMaxSave := 50.0, [5,12].EnableCfg := 1, [5,12].OverrideCfg := 1, [5,13].TagName := 'PI002', [5,13].OutofRange := 1, [5,13].Address := 13, [5,13].RawMin := 6553, [5,13].RawMax := 32767, [5,13].RawLowLimit := 6225, [5,13].RawHighLimit := 33095, [5,13].FilterActual := 1.0, [5,13].ScaledMax := 100.0, [5,13].CurrentValue := -24.998093, [5,13].RangeMax := 100.0, [5,13].RangeMaxSave := 100.0, [5,13].RealCfg := 1, [5,13].EnableCfg := 1, [5,13].OverrideCfg := 1, [5,14].OutofRange := 1, [5,14].Address := 14, [5,14].RawMin := 5529, [5,14].RawMax := 27648, [5,14].RawLowLimit := 5253, [5,14].RawHighLimit := 27924, [5,14].FilterActual := 1.0, [5,14].ScaledMax := 14.0, [5,14].RangeMax := 14.0, [5,14].RangeMaxSave := 14.0, [5,14].RealCfg := 1, [5,14].OverrideCfg := 1, [5,15].OutofRange := 1, [5,15].Address := 15, [5,15].RawMin := 5529, [5,15].RawMax := 27648, [5,15].RawLowLimit := 5253, [5,15].RawHighLimit := 27924, [5,15].FilterActual := 1.0, [5,15].ScaledMax := 2.0, [5,15].CurrentValue := -0.49993217,
        [5,15].RangeMax := 2.0, [5,15].RangeMaxSave := 2.0, [5,15].RealCfg := 1, [5,15].OverrideCfg := 1, [5,16].OutofRange := 1, [5,16].Address := 16, [5,16].RawMin := 5529, [5,16].RawMax := 27648, [5,16].RawLowLimit := 5253, [5,16].RawHighLimit := 27924, [5,16].FilterActual := 1.0, [5,16].ScaledMax := 2.0, [5,16].CurrentValue := -0.49993217, [5,16].RangeMax := 2.0, [5,16].RangeMaxSave := 2.0, [5,16].RealCfg := 1, [5,16].OverrideCfg := 1, [5,17].OutofRange := 1, [5,17].Address := 17, [5,17].RawMin := 5529, [5,17].RawMax := 27648, [5,17].RawLowLimit := 5253, [5,17].RawHighLimit := 27924, [5,17].FilterActual := 1.0, [5,17].ScaledMin := -1.0, [5,17].ScaledMax := 5.0, [5,17].CurrentValue := -2.4997964, [5,17].RangeMin := -1.0, [5,17].RangeMax := 5.0, [5,17].RangeMinSave := -1.0, [5,17].RangeMaxSave := 5.0, [5,17].RealCfg := 1, [5,17].OverrideCfg := 1, [5,18].OutofRange := 1, [5,18].Address := 18, [5,18].RawMin := 5529, [5,18].RawMax := 27648, [5,18].RawLowLimit := 5253, [5,18].RawHighLimit := 27924, [5,18].FilterActual := 1.0, [5,18].ScaledMin := -1.0, [5,18].ScaledMax := 5.0, [5,18].CurrentValue := -2.4997964, [5,18].RangeMin := -1.0, [5,18].RangeMax := 5.0, [5,18].RangeMinSave := -1.0, [5,18].RangeMaxSave := 5.0, [5,18].RealCfg := 1, [5,18].OverrideCfg := 1, [5,19].OutofRange := 1, [5,19].Address := 19, [5,19].RawMin := 5529, [5,19].RawMax := 27648, [5,19].RawLowLimit := 5253, [5,19].RawHighLimit := 27924, [5,19].FilterActual := 1.0, [5,19].ScaledMin := -1.0, [5,19].ScaledMax := 5.0, [5,19].CurrentValue := -2.4997964, [5,19].RangeMin := -1.0,
        [5,19].RangeMax := 5.0, [5,19].RangeMinSave := -1.0, [5,19].RangeMaxSave := 5.0, [5,19].RealCfg := 1, [5,19].OverrideCfg := 1, [5,20].OutofRange := 1, [5,20].Address := 20, [5,20].RawMin := 5529, [5,20].RawMax := 27648, [5,20].RawLowLimit := 5253, [5,20].RawHighLimit := 27924, [5,20].FilterActual := 1.0, [5,20].ScaledMax := 100.0, [5,20].CurrentValue := -24.996607, [5,20].RangeMax := 100.0, [5,20].RangeMaxSave := 100.0, [5,20].RealCfg := 1, [5,20].OverrideCfg := 1, [5,21].OutofRange := 1, [5,21].Address := 21, [5,21].RawMin := 5529, [5,21].RawMax := 27648, [5,21].RawLowLimit := 5253, [5,21].RawHighLimit := 27924, [5,21].FilterActual := 1.0, [5,21].ScaledMax := 100.0, [5,21].CurrentValue := -24.996607, [5,21].RangeMax := 100.0, [5,21].RangeMaxSave := 100.0, [5,21].RealCfg := 1, [5,21].OverrideCfg := 1, [5,22].TagName := 'SPARE', [5,22].Address := 22, [5,22].RawMin := 5529, [5,22].RawMax := 27648, [5,22].RealCfg := 1, [5,22].OverrideCfg := 1, [5,23].TagName := 'SPARE', [5,23].Address := 23, [5,23].RawMin := 5529, [5,23].RawMax := 27648, [5,23].RealCfg := 1, [5,23].OverrideCfg := 1, [5,24].TagName := 'SPARE', [5,24].Address := 24, [5,24].RawMin := 5529, [5,24].RawMax := 27648, [5,24].RealCfg := 1, [5,24].OverrideCfg := 1, [5,25].TagName := 'SPARE', [5,25].Address := 25, [5,25].RawMin := 5529, [5,25].RawMax := 27648, [5,25].RealCfg := 1, [5,25].OverrideCfg := 1, [5,26].TagName := 'SPARE', [5,26].Address := 26, [5,26].RawMin := 5529, [5,26].RawMax := 27648, [5,26].RealCfg := 1,
        [5,26].OverrideCfg := 1, [5,27].TagName := 'SPARE', [5,27].Address := 27, [5,27].RawMin := 5529, [5,27].RawMax := 27648, [5,27].RealCfg := 1, [5,27].OverrideCfg := 1, [5,28].TagName := 'AI#1', [5,28].OutofRange := 1, [5,28].Address := 28, [5,28].RawMin := 6553, [5,28].RawMax := 32767, [5,28].RawLowLimit := 6225, [5,28].RawHighLimit := 33095, [5,28].FilterActual := 1.0, [5,28].ScaledMax := 100.0, [5,28].CurrentValue := -24.998093, [5,28].RangeMax := 100.0, [5,28].RangeMaxSave := 100.0, [5,28].RealCfg := 1, [5,28].EnableCfg := 1, [5,28].OverrideCfg := 1, [5,29].TagName := 'AI#2', [5,29].OutofRange := 1, [5,29].Address := 29, [5,29].RawMin := 6553, [5,29].RawMax := 32767, [5,29].RawLowLimit := 6225, [5,29].RawHighLimit := 33095, [5,29].FilterActual := 1.0, [5,29].ScaledMax := 100.0, [5,29].CurrentValue := -24.998093, [5,29].RangeMax := 100.0, [5,29].RangeMaxSave := 100.0, [5,29].RealCfg := 1, [5,29].EnableCfg := 1, [5,29].OverrideCfg := 1, [5,30].TagName := 'AI#3', [5,30].OutofRange := 1, [5,30].Address := 30, [5,30].RawMin := 6553, [5,30].RawMax := 32767, [5,30].RawLowLimit := 6225, [5,30].RawHighLimit := 33095, [5,30].FilterActual := 1.0, [5,30].ScaledMax := 100.0, [5,30].CurrentValue := -24.998093, [5,30].RangeMax := 100.0, [5,30].RangeMaxSave := 100.0, [5,30].RealCfg := 1, [5,30].EnableCfg := 1, [5,30].OverrideCfg := 1, [5,31].TagName := 'AI#4', [5,31].OutofRange := 1, [5,31].Address := 31, [5,31].RawMin := 6553, [5,31].RawMax := 32767, [5,31].RawLowLimit := 6225, [5,31].RawHighLimit := 33095, [5,31].FilterActual := 1.0,
        [5,31].ScaledMax := 100.0, [5,31].CurrentValue := -24.998093, [5,31].RangeMax := 100.0, [5,31].RangeMaxSave := 100.0, [5,31].RealCfg := 1, [5,31].EnableCfg := 1, [5,31].OverrideCfg := 1, [5,40].TagName := 'FI003', [5,40].Address := 40, [5,40].RawMin := 5529, [5,40].RawMax := 27648, [5,40].RawLowLimit := 5253, [5,40].RawHighLimit := 27924, [5,40].FilterActual := 1.0, [5,40].ScaledMax := 50.0, [5,40].RangeMax := 50.0, [5,40].RangeMaxSave := 50.0, [5,40].EnableCfg := 1, [5,40].OverrideCfg := 1, [5,41].TagName := 'LV003', [5,41].Address := 41, [5,41].RawMin := 6553, [5,41].RawMax := 32767, [5,41].RawLowLimit := 6225, [5,41].RawHighLimit := 33095, [5,41].FilterActual := 1.0, [5,41].ScaledMax := 99999.0, [5,41].RangeMax := 99999.0, [5,41].RangeMaxSave := 99999.0, [5,41].EnableCfg := 1, [5,41].OverrideCfg := 1, [5,42].TagName := 'LV001', [5,42].Address := 42, [5,42].RawMin := 6553, [5,42].RawMax := 32767, [5,42].RawLowLimit := 6225, [5,42].RawHighLimit := 33095, [5,42].FilterActual := 1.0, [5,42].ScaledMin := -1.0, [5,42].ScaledMax := 5.0, [5,42].RangeMin := -1.0, [5,42].RangeMax := 5.0, [5,42].RangeMinSave := -1.0, [5,42].RangeMaxSave := 5.0, [5,42].EnableCfg := 1, [5,42].OverrideCfg := 1, [5,43].TagName := 'LV002', [5,43].Address := 43, [5,43].RawMin := 6553, [5,43].RawMax := 32767, [5,43].RawLowLimit := 6225, [5,43].RawHighLimit := 33095, [5,43].FilterActual := 1.0, [5,43].ScaledMax := 99999.0, [5,43].RangeMax := 99999.0, [5,43].RangeMaxSave := 99999.0, [5,43].EnableCfg := 1, [5,43].OverrideCfg := 1, [5,44].Address := 44, [5,44].RawMin := 6553,
        [5,44].RawMax := 32767, [5,44].RawLowLimit := 6225, [5,44].RawHighLimit := 33095, [5,44].FilterActual := 1.0, [5,44].ScaledMax := 99999.0, [5,44].RangeMax := 99999.0, [5,44].RangeMaxSave := 99999.0, [5,45].Address := 42, [5,45].RawMin := 6553, [5,45].RawMax := 32767, [5,45].RawLowLimit := 6225, [5,45].RawHighLimit := 33095, [5,45].FilterActual := 1.0, [5,45].ScaledMin := -1.0, [5,45].ScaledMax := 5.0, [5,45].RangeMin := -1.0, [5,45].RangeMax := 5.0, [5,45].RangeMinSave := -1.0, [5,45].RangeMaxSave := 5.0, [5,45].OverrideCfg := 1);
   AO1 : ALIAS FOR AnalogOutput[8];
   AO2 : ALIAS FOR AnalogOutput[9];
   AO3 : ALIAS FOR AnalogOutput[10];
   AO4 : ALIAS FOR AnalogOutput[11];
   AP008 : ALIAS FOR DigitalOutput[14];
   ARC_AI101 : ARC_pH := (ProductAssignTime := 1743405110, W_CALIBVALUES_Offset := 7.0, W_CALIBVALUES_Slope := -58.92, W_CALIBVALUES_Temp := 298.15, W_CALIBPROD_Command := 1, W_CALIBPRODVAL_Value := 7.0, W_SYNCTIME_Time := 1759491692, W_USER_Level := 48, W_USER_Password := 16021966);
   ARC_AI202 : ARC_pH := (ProductAssignTime := 1727190388, W_CALIBVALUES_Offset := 3.0, W_CALIBVALUES_Slope := -58.21, W_CALIBVALUES_Temp := 298.15, W_CALIBPROD_Command := 1, W_CALIBPRODVAL_Value := 7.0, W_SYNCTIME_Time := 1759491693, W_USER_Level := 48, W_USER_Password := 16021966);
   BagInflate : BagInflate := (SP := 10.0, PV := -34.497368);
   BAN001P : ALIAS FOR DigitalOutput[4];
   BAN001S : ALIAS FOR DigitalOutput[3];
   BAN002P : ALIAS FOR DigitalOutput[6];
   BAN002S : ALIAS FOR DigitalOutput[5];
   CCPSystem : CCPSystem := (Download := 1, OperationDownloadFlag := 1, Manual := 1, State := 3, Language := 1, EndPointer := 81, Machine := 'Mobius TFF', Created := '01/31/2025 6:03:13 PM', Originator := 'Joshua korba', OperationName := 'c:\\Smart\\TFF80\\CCPRecipeFiles\\W2882\\W2882 2200 - 3200g UFDF_01.00.opn', ConfigFile := 'RDP2306026_TFF80.cfg', StateWatchDog.PRE := 300000, EventList.Event[0] := 709, EventList.Event[1] := 600101, EventList.Event[2] := 2500101, EventList.Event[3] := 2500301, EventList.Event[4] := 2500401, EventList.Event[5] := 2500501, EventList.Event[6] := 2500601, EventList.Event[7] := 2500701, EventList.Event[8] := 2500801, EventList.Event[9] := 2500901, EventList.Event[10] := 2501001, EventList.Event[11] := 2501101, EventList.Event[12] := 2501201, EventList.Event[13] := 2501301, EventList.Event[14] := 2501401, EventList.Event[15] := 2501501, EventList.Event[16] := 2501601, EventList.Event[17] := 2501701, EventList.Event[18] := 2501801, EventList.Event[19] := 2501901, EventList.Event[20] := 2502001, EventList.Event[21] := 2502101, EventList.Event[22] := 2502201, EventList.Event[23] := 2502801, EventList.Event[24] := 2502901, EventList.Event[25] := 2503001, EventList.Event[26] := 2503101, EventList.Event[27] := 2503201, EventList.Event[28] := 2503301, EventList.Event[29] := 2504001, EventList.Event[30] := 2504101, EventList.Event[31] := 2504201, EventList.Event[32] := 2504301, EventList.Event[33] := 2504401, EventList.Event[34] := 1300001, EventList.Event[35] := 1300101, EventList.Event[36] := 1300201, EventList.Event[37] := 1300301, EventList.Event[38] := 1300401, EventList.Event[39] := 1300501, EventList.Event[40] := 1300601, EventList.Event[41] := 1300701, EventList.Event[42] := 1300801, EventList.Event[43] := 1300901, EventList.Event[44] := 1301001, EventList.Event[45] := 1301101, EventList.Event[46] := 1301201, EventList.Event[47] := 1301501,
        EventList.Event[48] := 1301601, EventList.Event[49] := 1301701, EventList.Event[50] := 1301801, EventList.Event[51] := 1301901, EventList.Event[52] := 1302001, EventList.Event[53] := 2600001, EventList.Event[54] := 2600002, EventList.Event[55] := 2600003, EventList.Event[56] := 2600004, EventList.Event[57] := 900101, EventList.Event[58] := 500101, EventList.Event[59] := 500102, EventList.Event[60] := 500103, EventList.Event[61] := 500104, EventList.Event[62] := 500106, EventList.Event[63] := 500107, EventList.Event[64] := 500108, EventList.Event[65] := 500109, EventList.Event[66] := 500111, EventList.Event[67] := 500112, EventList.Event[68] := 500113, EventList.Event[69] := 500114, EventList.Event[70] := 500115, EventList.Event[71] := 500116, EventList.Event[72] := 500117, EventList.Event[73] := 500118, EventList.Event[74] := 500119, EventList.Event[75] := 500120, EventList.Event[76] := 500121, EventList.Event[77] := 500122, EventList.Event[78] := 500123, EventList.Event[79] := 500124, EventList.Event[80] := 500125, EventList.Event[81] := 200101, EventList.Event[82] := 200104, EventList.Event[83] := 200105, EventList.Event[84] := 900201, EventList.Event[85] := 500201, EventList.Event[86] := 500202, EventList.Event[87] := 500203, EventList.Event[88] := 500206, EventList.Event[89] := 500207, EventList.Event[90] := 500208, EventList.Event[91] := 500211, EventList.Event[92] := 500212, EventList.Event[93] := 500213, EventList.Event[94] := 500214, EventList.Event[95] := 500215, EventList.Event[96] := 500216, EventList.Event[97] := 500217, EventList.Event[98] := 500218, EventList.Event[99] := 500219, EventList.Event[100] := 500220, EventList.Event[101] := 500221, EventList.Event[102] := 200201, EventList.Event[103] := 200204, EventList.Event[104] := 200205, EventList.Event[105] := 900301, EventList.Event[106] := 1400001, EventList.Event[107] := 1400002,
